(* IEC 61131-3 sources: daoli-st-library/DL_Process (part 27) *)

(* ---- FB_DL_ChillerCondReset.st ---- *)
(*
  FB_DL_ChillerCondReset  —  冷水机组冷凝压力重置（室外湿球联动限幅） / Chiller condensing-pressure setpoint reset driven by outdoor wet-bulb with clamping
  分类 Category : DL_Process
  版本 Version  : 1.0.0
  来源 Source   : t1-2-oscat-building — 楼宇冷站冷凝压力重置族深化
  溯源 Origin   : 道莅 clean-room 实现；湿球联动线性重置 + 死区 + 步长限幅为公开 HVAC 节能控制律，未复制任何源码行
  功能 Function : 1) 目标设定 fCondSpKpa = fWetBulbC × fSlopeKpaPerK + fOffsetKpa；
                  2) 硬限幅钳制到 [fSpMinKpa, fSpMaxKpa]（先限幅后限速，顺序固定）；
                  3) 步长限速：单次调用变化量不超过 fStepMaxKpa（向上与向下同限）；
                  4) 死区保持：|候选 - 当前输出| < fDeadbandKpa 时输出保持不变（避免阀位抖动）；
                  5) 故障级单码 03A3，归因由 eCause 独立成员承载（R190）；
                  6) 信息级 04CB = 重置激活沿（进 eRun 单拍）；7) 解除式全当拍量（R240）。
  接口 Interface: 输入湿球/斜率/偏置/上下限/死区/步长；输出设定值与限幅/限速镜像
  边界 Boundary : ① 组态闸：fSlopeKpaPerK <= 0.0、fSpMaxKpa <= fSpMinKpa、fStepMaxKpa <= 0.0、
                  fDeadbandKpa < 0.0、fWetBulbMaxC <= fWetBulbMinC 任一成立 → 03A3 锁存；
                  ② 湿球非有限（NaN 自反 + Inf 差值自减）或越量程 → 03A3 锁存，输出保持上一有效值
                  （冻结保持，非降级）；③ 浮点判据全容差式，禁 = / <> 判等；
                  ④ 无 TON 跨相复用（仅一个激活沿 R_TRIG + 一个 R_TRIG 复位沿），段 0 无条件调用；
                  ⑤ 故障相迁出唯一路径 = bReset 上升沿；⑥ 零全局耦合（无 GVL / %I %Q %M）。
  依赖 Depends  : Standard.library（R_TRIG）
  码表 Error codes（Process 段 0005，故障窗口 03A3 / 信息窗口 04CB）:
    16#0005_03A3 故障级：冷凝压力重置故障总码（组态非法 / 湿球非有限 / 湿球越量程），
                 锁存至 bReset 上升沿；归因见 eCause，不新增码位（派单硬约束单码）
    16#0005_04CB 信息级：重置激活沿（bEnable 上升进入 eRun 单拍）
  修订历史 Revision :
    2026-11-19  v1.0.0  R43 首版（批次 2 · 序号 7）
*)

TYPE E_DL_CcrState :
(
    eIdle  := 0,      // 未使能：输出冻结上一值 / Idle, output frozen
    eRun   := 10,     // 重置运行中 / Reset active
    eFault := 90      // 故障锁存相 / Fault latched phase
);
END_TYPE

TYPE E_DL_CcrCause :
(
    eNone       := 0, // 无故障成因 / No cause
    eCfgIllegal := 1, // 组态非法 / Illegal configuration
    eWbNonFin   := 2, // 湿球输入非有限 / Wet-bulb non-finite
    eWbRange    := 3  // 湿球越量程 / Wet-bulb out of range
);
END_TYPE

FUNCTION_BLOCK FB_DL_ChillerCondReset
VAR_INPUT
    fWetBulbC      : REAL := 10.0;     // 室外湿球温度 [°C] / Outdoor wet-bulb temperature
    fWetBulbMinC   : REAL := -20.0;    // 湿球量程下限 [°C] / Wet-bulb range low
    fWetBulbMaxC   : REAL := 45.0;     // 湿球量程上限 [°C] / Wet-bulb range high
    fSlopeKpaPerK  : REAL := 2.0;      // 联动斜率 [kPa/K]，域 > 0 / Reset slope
    fOffsetKpa     : REAL := 400.0;    // 联动偏置 [kPa] / Reset offset
    fSpMinKpa      : REAL := 500.0;    // 设定下限 [kPa] / Setpoint low limit
    fSpMaxKpa      : REAL := 900.0;    // 设定上限 [kPa] / Setpoint high limit
    fDeadbandKpa   : REAL := 5.0;      // 死区 [kPa]，域 >= 0 / Deadband
    fStepMaxKpa    : REAL := 10.0;     // 单次限速步长 [kPa]，域 > 0 / Rate limit step
    bEnable        : BOOL := FALSE;    // 重置使能（电平）[-] / Reset enable
    bReset         : BOOL := FALSE;    // 复位命令，上升沿清故障 [-] / Reset edge
END_VAR
VAR_OUTPUT
    eState         : E_DL_CcrState;    // 状态出口，段 6 单点映射 / State outlet
    eCause         : E_DL_CcrCause;    // 故障成因出口（R190） / Fault cause outlet
    fCondSpKpa     : REAL;             // 冷凝压力设定 [kPa] / Condensing pressure setpoint
    bLimited       : BOOL;             // 限幅生效镜像 [-] / Clamp active mirror
    bDbHold        : BOOL;             // 死区保持镜像 [-] / Deadband hold mirror
    bError         : BOOL;             // 故障锁存标志 [-] / Fault latch flag
    nErrId         : UDINT;            // 事件码，0 = 无事件 / Event code
END_VAR
VAR
    _eState        : E_DL_CcrState := E_DL_CcrState.eIdle;   // 内部相位（CASE 唯一写入目标） / Internal phase
    _eCause        : E_DL_CcrCause := E_DL_CcrCause.eNone;   // 故障成因锁存（锁存量） / Latched cause
    rtEnable       : R_TRIG;           // 使能沿实例，每周期无条件调用 / Enable edge
    rtReset        : R_TRIG;           // 复位沿实例，每周期无条件调用 / Reset edge
    _fSp           : REAL;             // 设定输出保持槽（持久） / Setpoint holding slot
    _fRawKpa       : REAL;             // 未限幅原始设定 [kPa]（当拍量） / Raw setpoint
    _fClampKpa     : REAL;             // 限幅后候选 [kPa]（当拍量） / Clamped candidate
    _bClampOn      : BOOL;             // 限幅生效当拍量 [-] / Clamp active
    _bNonFin       : BOOL;             // 湿球非有限当拍量 [-] / Wet-bulb non-finite
    _bRangeBad     : BOOL;             // 湿球越量程当拍量 [-] / Wet-bulb out of range
    _bCfgBad       : BOOL;             // 组态非法当拍量 [-] / Config illegal
    _bFault        : BOOL;             // 故障锁存位（锁存量） / Latched fault bit
    _uFault        : UDINT;            // 故障码锁存（锁存量） / Latched fault code
    _uInfo         : UDINT;            // 信息码，每拍重算 / Transient info code
END_VAR

(* —— 段 0：沿实例无条件周期刷新 + 当拍量判据 —— *)
_fRawKpa := fWetBulbC * fSlopeKpaPerK + fOffsetKpa;                       // 联动原始设定 [kPa] / Raw linked setpoint
_bNonFin := (fWetBulbC <> fWetBulbC) OR ((fWetBulbC - fWetBulbC) <> (fWetBulbC - fWetBulbC));   // NaN/Inf 双判 / NaN and Inf
_bRangeBad := (fWetBulbC < fWetBulbMinC) OR (fWetBulbC > fWetBulbMaxC);    // 量程判据（双侧直比） / Range verdict
_bCfgBad := (fSlopeKpaPerK <= 0.0) OR (fSpMaxKpa <= fSpMinKpa) OR (fStepMaxKpa <= 0.0)
            OR (fDeadbandKpa < 0.0) OR (fWetBulbMaxC <= fWetBulbMinC);     // 组态非法当拍量 / Config illegal
rtEnable(CLK := bEnable);                                                 // 使能沿，每拍必调 / Enable edge
rtReset(CLK := bReset);                                                   // 复位沿，每拍必调 / Reset edge

(* —— 段 1：单拍量预清零（锁存量与设定保持槽不入清单） —— *)
_uInfo := 16#0000_0000;            // 信息码每拍重算 / Info recomputed
bLimited := FALSE;                 // 限幅镜像缺省 FALSE / Clamp mirror default
bDbHold := FALSE;                  // 死区镜像缺省 FALSE / Deadband mirror default
nErrId := 16#0000_0000;            // 事件码缺省无事件 / Event code default

(* —— 段 2：复位沿 + 组态域闸 —— *)
IF rtReset.Q THEN                              // rtReset.Q = 当拍量 / current scan
    _bFault := FALSE;                          // 清故障锁存位（锁存量） / Clear fault latch
    _uFault := 16#0000_0000;                   // 清故障锁存码（锁存量） / Clear fault code
    _eCause := E_DL_CcrCause.eNone;            // 清成因（锁存量） / Clear cause
    IF _eState = E_DL_CcrState.eFault THEN
        _eState := E_DL_CcrState.eIdle;        // 故障相迁出：回未使能 / Fault exit to idle
    END_IF
END_IF
IF _bCfgBad THEN                               // 组态域闸 / Config gate
    _uFault := 16#0005_03A3;                   // 故障级：重置故障总码 / Process fault code
    _eCause := E_DL_CcrCause.eCfgIllegal;      // 归因：组态非法 / Cause: illegal config
    _bFault := TRUE;                           // 标志与码位配对（R45） / Flag paired with code
END_IF

(* —— 段 3：湿球非有限 / 越量程（判据当拍量） —— *)
IF (NOT _bFault) AND _bNonFin THEN             // 非有限锁存 / Non-finite latch
    _uFault := 16#0005_03A3;
    _eCause := E_DL_CcrCause.eWbNonFin;        // 归因：非有限 / Cause: non-finite
    _bFault := TRUE;
END_IF
IF (NOT _bFault) AND (NOT _bNonFin) AND _bRangeBad THEN   // 越量程锁存 / Range latch
    _uFault := 16#0005_03A3;
    _eCause := E_DL_CcrCause.eWbRange;         // 归因：越量程 / Cause: out of range
    _bFault := TRUE;
END_IF

(* —— 段 4：故障解除式（R240；全当拍量）：rtReset.Q / NOT _bCfgBad / NOT _bNonFin / NOT _bRangeBad —— *)
IF rtReset.Q AND (NOT _bCfgBad) AND (NOT _bNonFin) AND (NOT _bRangeBad) THEN
    _bFault := FALSE;                          // 清故障锁存位（锁存量） / Clear fault latch
    _uFault := 16#0000_0000;                   // 清故障锁存码（锁存量） / Clear fault code
    _eCause := E_DL_CcrCause.eNone;            // 清成因（锁存量） / Clear cause
END_IF

(* —— 段 4A：故障锁存相位迁移闸（输出冻结上一有效值，非降级） —— *)
IF _bFault AND (_eState <> E_DL_CcrState.eFault) THEN
    _eState := E_DL_CcrState.eFault;           // 锁存即入故障相 / Latch enters fault phase
END_IF

(* —— 段 5：相位机（CASE 全覆盖 + ELSE 兜底） —— *)
CASE _eState OF

E_DL_CcrState.eIdle:
    IF rtEnable.Q AND (NOT _bFault) THEN       // 使能上升沿启动 / Enable rising starts
        _uInfo := 16#0005_04CB;                // 信息级：重置激活沿 / Info: reset active edge
        _eState := E_DL_CcrState.eRun;         // 进运行相 / Enter run
    END_IF

E_DL_CcrState.eRun:
    IF NOT bEnable THEN                        // 撤使能：回未使能（输出冻结） / Disable returns idle
        _eState := E_DL_CcrState.eIdle;
    ELSE
        _fClampKpa := _fRawKpa;                            // 候选 = 原始设定 / Candidate from raw
        IF _fClampKpa < fSpMinKpa THEN                     // 下限钳制 / Low clamp
            _fClampKpa := fSpMinKpa;
            _bClampOn := TRUE;
        ELSIF _fClampKpa > fSpMaxKpa THEN                  // 上限钳制 / High clamp
            _fClampKpa := fSpMaxKpa;
            _bClampOn := TRUE;
        ELSE
            _bClampOn := FALSE;                            // 未限幅 / No clamp
        END_IF
        IF ABS(_fClampKpa - _fSp) < fDeadbandKpa THEN      // 死区内保持（容差式比较） / Deadband hold
            bDbHold := TRUE;
        ELSIF (_fClampKpa - _fSp) > fStepMaxKpa THEN       // 向上限速 / Upward rate limit
            _fSp := _fSp + fStepMaxKpa;
        ELSIF (_fSp - _fClampKpa) > fStepMaxKpa THEN       // 向下限速 / Downward rate limit
            _fSp := _fSp - fStepMaxKpa;
        ELSE
            _fSp := _fClampKpa;                            // 直接跟随 / Direct follow
        END_IF
        IF (_fSp < fSpMinKpa) THEN                         // 限速后二次下限复核 / Post-limit low check
            _fSp := fSpMinKpa;
        ELSIF (_fSp > fSpMaxKpa) THEN                      // 限速后二次上限复核 / Post-limit high check
            _fSp := fSpMaxKpa;
        END_IF
    END_IF

E_DL_CcrState.eFault:
    ;                                          // 故障相：输出冻结，仅段 4 复位沿可迁出 / Frozen, reset only

ELSE
    _uFault := 16#0005_03A3;                   // 故障级：非法相位兜底（归并总码） / Illegal phase fallback
    _eCause := E_DL_CcrCause.eCfgIllegal;      // 归因：相位非法归并组态 / Cause: phase illegal
    _bFault := TRUE;
    _eState := E_DL_CcrState.eFault;           // 强制回故障相 / Force fault phase

END_CASE

(* —— 段 6：出口单点映射（名实同源；锁存码回放） —— *)
fCondSpKpa := _fSp;                            // 设定值出口 / Setpoint outlet
bLimited := _bClampOn AND (NOT _bFault);       // 限幅镜像 / Clamp mirror
bDbHold := bDbHold AND (NOT _bFault);          // 死区保持镜像 / Deadband mirror
IF _bFault THEN
    nErrId := _uFault;                         // 故障锁存码回放 / Replay latched code
ELSE
    nErrId := _uInfo;                          // 信息码 / Transient info
END_IF
bError := _bFault;                             // 故障标志同源 / Flag from latch
eState := _eState;                             // 状态出口 / State outlet
eCause := _eCause;                             // 成因出口 / Cause outlet

END_FUNCTION_BLOCK

(* ---- FB_DL_ChillerDoorPurgeSeq.st ---- *)
(*
    FB_DL_ChillerDoorPurgeSeq —— 冷机检修门吹扫联锁时序
    ------------------------------------------------------------------
    分类      : DL_Process / Interlock
    前缀      : FB_DL_
    版本      : 1.0.0
    溯源      : clean-room 自有实现；仅借鉴「先吹扫置换、后放行开门」的受限空间
                进入公开安全常识语义，未复制任何闭源厂商源码，码位 100% 自有
    平台      : 纯 IEC 61131-3，CODESYS V3.5+ / TwinCAT 3 / InoProShop / Machine Expert 通用
    作者      : 道莅代码库 · PLC编程专家（R76 冲刺批 C3 · #3）
    ------------------------------------------------------------------
    功能说明  : 冷机检修门「吹扫联锁」唯一时序属主件：门关到位确认 → 风压建立确认
                （fAirPress > fPressMin 持续 tPressQual，超 tPressTo 未建立报 1F00）
                → 吹扫倒计时（tPurgeDur）→ 吹扫完成（bDone 单拍脉冲）→ 放行门开允许
                （bDoorPermit）。任一异常（门中途打开 / 风压跌落 / 确认超时）→
                回退安全态（吹扫输出与开门允许同时撤销）并锁存故障，须 bReset 复位；
                bEStop 急停为最高优先，任意态立即回安全态并锁存 1F03。
                边界：只产出吹扫输出与开门允许，不驱动门电机、不判冷剂浓度。
    序列      : eIdle --bDoorClosed--> ePressQual --fbPressQual.Q--> ePurging
                --fbPurge.Q--> eReady（bDoorPermit）--门正常打开--> eIdle；
                ePressQual/ePurging --门中途打开--> eFault（1F02）；
                ePurging --风压跌落--> eFault（1F01）；ePressQual --超时--> eFault（1F00）。
    错误码    : 16#0005_1F00 风压建立确认超时（tPressTo 内未持续达标）——故障级
                16#0005_1F01 吹扫期间风压跌落（低于 fPressMin）——故障级
                16#0005_1F02 门中途打开（风压确认或吹扫中）——故障级
                16#0005_1F03 急停触发——故障级，最高优先，任意态立即安全态
                16#0005_1F04 参数/采样非法（fAirPress 非有限 / 阈值非正 / 时间为零）——故障级
                16#0005_1F05 CASE 落 ELSE 兜底——故障级
    码位总账  : 16#0005_1F00..1F05 全部定义并使用，无空悬码位
    状态机    : E_DL_PurgeState（eIdle / ePressQual / ePurging / eReady / eFault），
                CASE 含 ELSE 兜底：落 ELSE 置 16#0005_1F05、回安全态转 eFault。
                全部故障码锁存至复位沿：bReset 上升沿且 bEStop 已解除方可复位；
                吹扫完成脉冲 bDone 为单拍位：内部 _bDonePulse 置位 → 统一出口
                映射单拍发布（两段式，防同拍抹除）。
    安全优先级: 段 3 急停拦截在参数门禁与状态机之前执行，任意态（含 eFault）急停
                即重锁存 1F03 并保持安全态输出；安全态 = 吹扫输出 OFF + 开门允许 OFF。
    定时器    : 三只 TON + 两只 R_TRIG 在本体段 1 无条件周期刷新（R7），绝不放入
                CASE/IF，实例无跨相复用。
    防御口径  : 浮点比较一律阈值比较（禁 =/<>）；本件无除法运算；非有限判定按
                NaN f<>f、±Inf (f-f)<>(f-f)。
    修订记录  : 2026-11-23 v1.0.0 首次入库（R76 冲刺批 C3 · #3）
*)
TYPE E_DL_PurgeState :
(
    eIdle       := 0,   // 待机，等门关到位，吹扫与放行全撤销 / idle, waiting for the closed door, purge and permit both off
    ePressQual  := 10,  // 风压建立确认中，fAirPress 持续达标计时 / pressure qualifying, timing while air pressure stays above the minimum
    ePurging    := 20,  // 吹扫倒计时中，风压须持续保持 / purging, countdown running while pressure must hold
    eReady      := 30,  // 吹扫完成，开门允许放行 / purge complete, door-open permit granted
    eFault      := 40   // 故障，安全态保持，故障码锁存至复位沿 / fault, safe state held, code latched until the reset edge
);
END_TYPE

FUNCTION_BLOCK FB_DL_ChillerDoorPurgeSeq
VAR_INPUT
    bDoorClosed : BOOL;                  // 门关到位反馈，TRUE = 已关严 / door closed feedback, TRUE = fully closed
    fAirPress   : REAL;                  // 吹扫风压采样 [kPa] / purge air pressure sample [kPa]
    fPressMin   : REAL := 5.0;           // 风压建立阈值 [kPa]，必须大于 0 / pressure qualification threshold [kPa], must exceed zero
    tPressQual  : TIME := T#1S;          // 风压确认持续时间 [ms]，必须大于 0 / pressure qualification dwell [ms], must exceed zero
    tPressTo    : TIME := T#5S;          // 风压建立超时窗 [ms]，须大于 tPressQual / pressure establish timeout [ms], must exceed tPressQual
    tPurgeDur   : TIME := T#30S;         // 吹扫倒计时时长 [ms]，必须大于 0 / purge duration [ms], must exceed zero
    bEStop      : BOOL;                  // 急停输入，TRUE = 急停，最高优先 / emergency stop, TRUE = stopped, highest priority
    bReset      : BOOL;                  // 故障复位请求，上升沿生效且须急停已解除 / fault reset request, edge-active and requires estop cleared
END_VAR
VAR_OUTPUT
    bPurgeCmd   : BOOL;                  // 吹扫风机/风阀输出，仅确认与吹扫相置位 / purge blower or valve output, asserted in the qualify and purge phases only
    bDoorPermit : BOOL;                  // 门开允许，仅吹扫完成相置位 / door-open permit, asserted in the ready phase only
    bDone       : BOOL;                  // 吹扫完成单拍脉冲，发布后自清 / purge-complete one-scan pulse, self-cleared after publishing
    eState      : E_DL_PurgeState;       // 当前状态镜像输出 / current state mirror output
    nErrCode    : UDINT;                 // 错误码，0 = 无错；故障级码全部锁存回放 / error code, 0 = none; all fault-class codes latched and replayed
    bError      : BOOL;                  // 故障级标志，仅故障级码置位 / fault-class flag, raised only by fault-class codes
    bValid      : BOOL;                  // 输出可用标志，= NOT bError / outputs valid flag, equals NOT bError
END_VAR
VAR
    fbPressQual : TON;                   // 风压确认定时器，仅 ePressQual 使用 / pressure qualification timer, ePressQual only
    fbPressTo   : TON;                   // 风压建立超时定时器，仅 ePressQual 使用 / pressure establish timeout timer, ePressQual only
    fbPurge     : TON;                   // 吹扫倒计时定时器，仅 ePurging 使用 / purge countdown timer, ePurging only
    rtReset     : R_TRIG;                // 复位上升沿检测 / reset rising-edge detector
    _eState     : E_DL_PurgeState;       // 当前状态 / current state
    _uErrLatch  : UDINT;                 // 故障码锁存副本，故障态每拍回放 / latched fault code republished inside the fault state
    _bDonePulse : BOOL;                  // 完成脉冲源，段 2 发布后立刻自清 / completion pulse source, published then cleared in segment 2
    _bGateOk    : BOOL;                  // 参数与采样门禁结果 / parameter and sample gate result
END_VAR
VAR CONSTANT
    DL_CDP_ZERO : REAL := 0.0;           // 零值常量，避免裸字面量 [kPa] / zero constant avoiding a bare literal [kPa]
    DL_CDP_T_ZERO : TIME := T#0S;        // 零时间常量，参数门禁用 / zero time constant for the parameter gate
END_VAR

// 段 1｜定时器与边缘检测无条件周期刷新（R7：严禁放入 IF / CASE，实例无跨相复用）
// segment 1, timers and edge detectors refreshed unconditionally, never inside IF/CASE, no cross-phase reuse
fbPressQual(IN := (_eState = E_DL_PurgeState.ePressQual) AND (fAirPress > fPressMin) AND _bGateOk, PT := tPressQual);
fbPressTo(IN := (_eState = E_DL_PurgeState.ePressQual), PT := tPressTo);
fbPurge(IN := (_eState = E_DL_PurgeState.ePurging), PT := tPurgeDur);
rtReset(CLK := bReset);

// 段 2｜输出与错误状态预置；故障态从锁存副本回放；完成脉冲统一出口单拍发布（两段式）
// segment 2, preset outputs and error status; the fault state replays from the latch; the done pulse is published one scan via the unified exit
bDone := _bDonePulse;                    // 发布上一拍置的完成脉冲 / publish the pulse latched last scan
_bDonePulse := FALSE;                    // 发布即自清，保证只出现一拍 / clear right after publishing so the pulse lasts one scan
nErrCode := 0;                           // 预置无错误码 / preset no error code
bError := FALSE;                         // 预置无故障标志 / preset no fault flag
bValid := TRUE;                          // 预置输出可用 / preset outputs valid
IF _eState = E_DL_PurgeState.eFault THEN
    nErrCode := _uErrLatch;              // 重发布锁存故障码，HMI 不会看到码位闪断 / republish the latched fault code
    bError := TRUE;                      // 故障态恒置故障标志 / fault flag stays raised in the fault state
    bValid := FALSE;                     // 故障态输出不可信 / outputs not valid in the fault state
END_IF

// 段 3｜急停最高优先拦截 + 参数/采样门禁：急停任意态立即锁存 1F03 回安全态；
//        门禁非法锁存 1F04 转故障；已在故障态不覆盖原锁存码
// segment 3, estop has the highest priority and latches 1F03 from any state including fault;
//        the parameter gate latches 1F04; an existing latch inside the fault state is not overwritten
IF bEStop THEN
    _uErrLatch := 16#0005_1F03;          // 锁存急停码（任意态含 eFault 均可覆盖更新）/ latch the estop code, overridable from any state
    nErrCode := 16#0005_1F03;            // 故障级码赋值 3 行内置 bError / fault-class assignment with bError inline
    bError := TRUE;
    bValid := FALSE;
    _eState := E_DL_PurgeState.eFault;   // 立即回安全态，本拍 CASE 按 eFault 分派 / jump to the safe state, CASE dispatches on eFault
ELSE
    _bGateOk := (fPressMin > DL_CDP_ZERO) AND (tPressQual > DL_CDP_T_ZERO)
            AND (tPressTo > DL_CDP_T_ZERO) AND (tPurgeDur > DL_CDP_T_ZERO)
            AND (tPressTo > tPressQual);
    IF (fAirPress <> fAirPress) OR ((fAirPress - fAirPress) <> (fAirPress - fAirPress)) THEN
        _bGateOk := FALSE;               // 风压采样 NaN 或 ±Inf，非有限判定 / pressure sample NaN or infinite
    END_IF
    IF (NOT _bGateOk) AND (_eState <> E_DL_PurgeState.eFault) THEN
        _uErrLatch := 16#0005_1F04;      // 锁存参数/采样非法码 / latch the illegal parameter or sample code
        nErrCode := 16#0005_1F04;        // 故障级码赋值 3 行内置 bError / fault-class assignment with bError inline
        bError := TRUE;
        bValid := FALSE;
        _eState := E_DL_PurgeState.eFault; // 参数不可信直接转故障 / untrusted parameters jump to fault
    END_IF
END_IF

// 段 4｜主状态机：CASE + ELSE 兜底（R6）；每个相注明 拍 N 进入 / 本拍行为 / 拍 N+1 转出
// segment 4, main state machine, CASE with ELSE fallback; each phase notes entry, per-scan behaviour and exits
CASE _eState OF
E_DL_PurgeState.eIdle:
    // 拍 N 进入：复位后或门正常打开后；本拍行为：全撤销等待；拍 N+1 转出：门关到位 → ePressQual
    // entered after reset or a normal door opening; everything off while waiting; exits to ePressQual on the closed door
    IF bDoorClosed AND _bGateOk THEN
        _eState := E_DL_PurgeState.ePressQual; // 进风压确认相，下一拍计时启动 / enter pressure qualification, timing starts next scan
    END_IF

E_DL_PurgeState.ePressQual:
    // 拍 N 进入：门关到位；本拍行为：风压达标则 fbPressQual 计时；拍 N+1 转出四路：
    // 计时到 → ePurging；门中途打开 → eFault（1F02）；确认超时 → eFault（1F00）；门禁 → eFault（段 3）
    // entered on the closed door; timer runs while pressure holds; exits to ePurging on Q,
    // to eFault on a mid-sequence door opening (1F02) or on the establish timeout (1F00)
    IF NOT bDoorClosed THEN
        _uErrLatch := 16#0005_1F02;      // 锁存门中途打开码 / latch the mid-sequence door opening code
        nErrCode := 16#0005_1F02;        // 故障级码赋值 3 行内置 bError / fault-class assignment with bError inline
        bError := TRUE;
        bValid := FALSE;
        _eState := E_DL_PurgeState.eFault; // 回安全态，吹扫与放行同拍撤销 / safe state, purge and permit drop the same scan
    ELSIF fbPressQual.Q THEN
        _eState := E_DL_PurgeState.ePurging; // 风压确认通过，进吹扫倒计时 / pressure qualified, start the purge countdown
    ELSIF fbPressTo.Q THEN
        _uErrLatch := 16#0005_1F00;      // 锁存风压建立超时码 / latch the pressure establish timeout code
        nErrCode := 16#0005_1F00;        // 故障级码赋值 3 行内置 bError / fault-class assignment with bError inline
        bError := TRUE;
        bValid := FALSE;
        _eState := E_DL_PurgeState.eFault; // 超时回退安全态 / roll back to the safe state on timeout
    END_IF

E_DL_PurgeState.ePurging:
    // 拍 N 进入：风压确认通过；本拍行为：吹扫输出保持、倒计时走、风压须持续达标；
    // 拍 N+1 转出三路：倒计时到 → eReady（置完成脉冲源）；风压跌落 → eFault（1F01）；
    // 门中途打开 → eFault（1F02）
    // entered after qualification; purge output held, countdown running, pressure must hold;
    // exits to eReady with the pulse source on Q, to eFault on pressure drop (1F01) or door opening (1F02)
    IF NOT bDoorClosed THEN
        _uErrLatch := 16#0005_1F02;      // 锁存门中途打开码 / latch the mid-sequence door opening code
        nErrCode := 16#0005_1F02;        // 故障级码赋值 3 行内置 bError / fault-class assignment with bError inline
        bError := TRUE;
        bValid := FALSE;
        _eState := E_DL_PurgeState.eFault; // 回安全态 / return to the safe state
    ELSIF fAirPress < fPressMin THEN
        _uErrLatch := 16#0005_1F01;      // 锁存风压跌落码 / latch the pressure drop code
        nErrCode := 16#0005_1F01;        // 故障级码赋值 3 行内置 bError / fault-class assignment with bError inline
        bError := TRUE;
        bValid := FALSE;
        _eState := E_DL_PurgeState.eFault; // 风压跌落立即回退 / roll back at once on the pressure drop
    ELSIF fbPurge.Q THEN
        _bDonePulse := TRUE;             // 置完成脉冲源，段 2 统一出口单拍发布 / set the pulse source, published one scan via segment 2
        _eState := E_DL_PurgeState.eReady;   // 吹扫完成，进放行相 / purge complete, enter the ready phase
    END_IF

E_DL_PurgeState.eReady:
    // 拍 N 进入：吹扫倒计时到；本拍行为：开门允许置位（输出映射段）、吹扫输出撤销；
    // 拍 N+1 转出：门正常打开（关反馈消失）→ eIdle，下次关门重新吹扫
    // entered when the countdown elapsed; permit asserted via the output map while the purge output drops;
    // exits to eIdle when the door actually opens, the next closure restarts the purge
    IF NOT bDoorClosed THEN
        _eState := E_DL_PurgeState.eIdle;    // 门已开，正常返回待机 / door opened, normal return to idle
    END_IF

E_DL_PurgeState.eFault:
    // 拍 N 进入：任一故障级路径；本拍行为：安全态保持、锁存码回放；拍 N+1 转出：
    // bReset 上升沿且急停已解除 → eIdle（门关反馈丢失自动回 eIdle 等下次关门）
    // entered from any fault path; safe state held and the latch replays; exits to eIdle only on
    // a reset edge with the estop cleared
    IF rtReset.Q AND (NOT bEStop) THEN
        _uErrLatch := 0;                 // 清锁存码 / clear the latched code
        _eState := E_DL_PurgeState.eIdle;    // 回待机，等下次门关到位 / back to idle for the next closure
    END_IF

ELSE
    // 非法状态拦截：任何未定义枚举值一律锁存兜底码并转故障（R6）
    // illegal-state interception, any undefined enum value latches the fallback code and goes to fault
    _uErrLatch := 16#0005_1F05;          // 锁存兜底码 / latch the fallback code
    nErrCode := 16#0005_1F05;            // 故障级码赋值 3 行内置 bError / fault-class assignment with bError inline
    bError := TRUE;
    bValid := FALSE;
    _eState := E_DL_PurgeState.eFault;
END_CASE

// 段 5｜输出映射：吹扫输出仅确认/吹扫相保持，开门允许仅就绪相置位，其余一律撤销（双保险）
// segment 5, output map; purge output held only in qualify/purge, permit only in ready, everything else dropped as a double cut
bPurgeCmd := (_eState = E_DL_PurgeState.ePressQual)
          OR (_eState = E_DL_PurgeState.ePurging);   // 吹扫输出按相映射 / purge output mapped by phase
bDoorPermit := (_eState = E_DL_PurgeState.eReady);   // 开门允许仅在放行相 / permit only in the ready phase
eState := _eState;                                   // 状态镜像输出 / state mirror output

END_FUNCTION_BLOCK

(* ---- FB_DL_ChillerLiftOptimize.st ---- *)
(*
  Component : FB_DL_ChillerLiftOptimize
  Category  : DL_Process
  Type      : FB
  Version   : 1.0.0
  CodeSeg   : 16#06_0_37
  Summary   : 冷机 Lift（冷凝-蒸发温差）优化限值：温差基线统计窗 + 设定值 RateLimiter 限速输出。
              Chiller lift optimization: condenser-evaporator baseline statistics window plus rate-limited setpoint.
  溯源声明  : 道莅自研 clean-room
  边界安全  : 温度非有限（NaN 自反 + Inf 上限）拦截；基线统计窗点数域闸（≥ 1）；
              统计窗未满时输出冻结在当前值并置 bBaselineReady=FALSE（按派单要点）；
              设定值输出过 RateLimiter 限速（每拍步进钳制，防设定值跳变）；全浮点比较带 fEps 容差。
  复用      : 无
*)

FUNCTION_BLOCK FB_DL_ChillerLiftOptimize
VAR_INPUT
    bRun        : BOOL;                 (* 优化使能 · Enable *)
    fCondTC     : LREAL;                (* 冷凝器温度 [degC] · Condenser temperature *)
    fEvapTC     : LREAL;                (* 蒸发器温度 [degC] · Evaporator temperature *)
    nWinScans   : INT := 600;           (* 基线统计窗长 [拍] · Baseline window length *)
    fStepMaxK   : LREAL := 0.1;         (* 设定值每拍最大步进 [K] · Setpoint max step per scan *)
    fDeadK      : LREAL := 0.5;         (* 优化死区 [K]，防频繁调节 · Optimization deadband *)
    fEps        : LREAL := 1.0E-6;      (* 浮点判零容差 [实数域] · Floating zero tolerance *)
END_VAR
VAR_OUTPUT
    fLiftNowK   : LREAL;                (* 当前 Lift [K] · Current lift *)
    fLiftBaseK  : LREAL;                (* 基线平均 Lift [K] · Baseline mean lift *)
    fSetK       : LREAL;                (* 优化设定值输出 [K]，已限速 · Rate-limited setpoint *)
    bBaselineReady: BOOL;               (* 基线窗满标志 · Baseline ready flag *)
    bError      : BOOL;                 (* 故障标志，与故障码配对 · Fault flag paired with codes *)
    uErrorId    : UDINT;                (* 事件码 16#0000_0037，0 无事件 · Event code *)
END_VAR
VAR
    uCode   : WORD;     (* 码位暂存，每拍重算 [码] · Code staging *)
    bSigOk  : BOOL;     (* 输入有效标志 · Input validity flag *)
    fSumK   : LREAL;    (* 窗内 Lift 累加和 [K·拍] · Window sum *)
    nFill   : INT;      (* 窗内已累计拍数 [拍] · Window filled scans *)
    fTargetK: LREAL;    (* 目标设定值 [K] · Target setpoint *)
    fStepK  : LREAL;    (* 本拍实际步进 [K] · Actual step this scan *)
    nCycles : UDINT;    (* 有效拍计数 [拍]，防回卷 · Valid scan count *)
END_VAR
VAR CONSTANT
    DL_CLO_WRAP : UDINT := 4294967290;  (* 计数防回卷余量 [拍] · Counter wrap guard *)
END_VAR

(* === 段 0 · 实例刷新 === *)
(* 无 TON/R_TRIG 实例：基线窗按拍计数；No timer instances, scan-counted window *)

(* === 段 1 · 输入校验与量程闸 === *)
uCode := 16#0000;                       // 每拍清码（可达清零基线）/ Clear codes each scan
bSigOk := (fCondTC = fCondTC) AND (fEvapTC = fEvapTC)               // 非有限拦截 / Non-finite guard
          AND (ABS(fCondTC) < 1.0E308) AND (ABS(fEvapTC) < 1.0E308) // Inf 上限判据 / Inf limit
          AND (nWinScans >= 1)                                      // 窗长域闸 / Window length gate
          AND (fStepMaxK > 0.0) AND (fDeadK >= 0.0);                // 步进正域闸 / Step and deadband gates
IF NOT bSigOk THEN
    uCode := 16#0037;                   // 故障级：域外，输出冻结 / Fault: domain invalid, frozen
END_IF

(* === 段 2 · 主逻辑：Lift 基线统计与设定值限速 === *)
IF bSigOk THEN
    fLiftNowK := fCondTC - fEvapTC;     (* 当前 Lift [K] / Current lift *)
    IF bRun THEN
        IF nFill < nWinScans THEN
            fSumK := fSumK + fLiftNowK; (* 窗内累加 / Accumulate in window *)
            nFill := nFill + 1;         (* 窗计数推进 / Advance the window count *)
            bBaselineReady := FALSE;    (* 窗未满：基线未就绪 / Window not full *)
        ELSE
            fLiftBaseK := fSumK / UDINT_TO_LREAL(INT_TO_UDINT(nWinScans));  (* 基线均值 [K] / Baseline mean *)
            bBaselineReady := TRUE;     (* 窗满：基线就绪 / Window full, baseline ready *)
            IF fLiftNowK > (fLiftBaseK + fDeadK) THEN
                fTargetK := fLiftBaseK; (* 超死区回基线目标 / Target back to baseline *)
            ELSE
                fTargetK := fSetK;      (* 死区内保持现值 / Hold inside the deadband *)
            END_IF
        END_IF
    ELSE
        nFill := 0;                     (* 撤使能重开统计窗 / Restart the window on disable *)
        fSumK := 0.0;
        bBaselineReady := FALSE;        (* 撤使能基线失效 / Baseline not ready *)
    END_IF
    (* RateLimiter：设定值每拍步进钳制 / Rate limiter: clamp the per-scan step *)
    fStepK := fTargetK - fSetK;         (* 目标差 [K] / Gap to target *)
    IF fStepK > fStepMaxK THEN
        fSetK := fSetK + fStepMaxK;     (* 正向限速 / Positive rate limit *)
    ELSIF fStepK < (-fStepMaxK) THEN
        fSetK := fSetK - fStepMaxK;     (* 负向限速 / Negative rate limit *)
    ELSE
        fSetK := fTargetK;              (* 一步到位 / Settle to target *)
    END_IF
END_IF

(* === 段 3 · 输出映射与故障码 === *)
IF bSigOk THEN
    IF nCycles < DL_CLO_WRAP THEN
        nCycles := nCycles + 1;         (* 有效拍计数 / Count valid scans *)
    END_IF
END_IF
bError := (uCode <> 16#0000);           (* 故障标志配对 / Fault flag paired *)
uErrorId := WORD_TO_UDINT(uCode);       (* 码位单点写入（16#0000_0037 形态）/ Single write point *)
END_FUNCTION_BLOCK

(* ---- FB_DL_ChillerSeqMgr.st ---- *)
//==============================================================================
// 功能块：FB_DL_ChillerSeqMgr ｜ 中文名称：冷水机组群控调度
// 所属子库：DL_Process ｜ 版本：v1.0.0 ｜ 兼容：CODESYS V3.5+ / TwinCAT 3 / 汇川 InoProShop
// 功能描述：6 台冷水机组群控：按平滑后负荷率加减机（加/减各带独立延迟，双延迟防抖动）
//           + 主备轮值均衡（委托 FB_DL_DutyStandbyRotation，最短运行/最短停机时长逻辑
//           一律由该件承担，本件只把 tMinRun/tMinStop 转发，绝不重复实现）+ 故障切备
//           （故障台由轮值件跳过）+ 供水低温保护（强制减机，防冻管）。本件不内联机组建模
//           与机组自身控制（压缩机/冷却水阀/防冻判据归设备层），只出启停命令与调度诊断。
// 开源溯源 (Origin)：道莅原创实现（参考 公开工程惯例 分类与参数域）
// 单位表：温度[摄氏度] / 负荷率与阈值[百分数] / 延迟与最小时长[min] / 扫描间隔[ms] /
//         台数[台] / 机组号[号]
// 错误码表：16#0005_040C 信息级（加/减机延迟计时中，尚未动作，不置 bError）/
//           16#0005_040D 信息级（供水温度低限保护强制减机，信息级不锁故障但强制动作）/
//           16#0005_0354 故障级（无可用机组：全故障或全不就绪，工艺停机级，置 bError）/
//           16#0005_0355 故障级（负荷率/阈值组态非法：减机阈值 ≥ 加机阈值、阈值越
//           0~100、台数组态非法；兼轮值件参数冲突透传——轮值件 bError 透传复位且只在
//           故障相处置，R115）/ 16#0005_0356 故障级（输入非有限独立分支显式映射入本槽，
//           兼状态机 ELSE 非法状态兜底）。0356 共用反证句：非有限与非法状态在现有输出
//           组合下不可观测出差异（均为 bError + 全撤指令 + bValid 撤 + eState 进 eFault），
//           §3 未给本件独立非有限槽，故显式复用不越段。
// 状态机：E_DL_ChillerGroupState（eIdle=0 待机 / eRunning=10 稳态调度 /
//           eStageUp=20 加机延迟中 / eStageDown=30 减机延迟中 / eLowSupply=40 供水低温
//           保护 / eFault=99 故障兜底），CASE 含 ELSE 兜底，ELSE 置 0356 且全撤指令。
// 边界行为：① 无可用机组（全故障或全不就绪）→ 故障 0354 + bNoAvailable（工艺停机级，
//           非提示级）；② 阈值组态非法（减机阈值 ≥ 加机阈值、阈值不在 0~100）→ 故障
//           0355；③ 供水温度 < fSupplyLowC → 强制减机一台 + 信息 040D + bLowSupplyProtect
//           （防冻管，信息级不锁故障但强制动作）；④ 加减机延迟计时中 → 信息 040C；
//           ⑤ 需求台数域 0~6 钳位，且不超过可用台数；⑥ 非有限 → 独立分支显式置 0356，
//           全撤指令；⑦ 失能 → 全撤指令 + bValid := FALSE（R72）；⑧ 轮值调用
//           FB_DL_DutyStandbyRotation（组合调用），tMinRunTime/tMinStopTime 由本件引脚
//           转发，最短运行/停机逻辑不重复实现；轮值件 bError 透传复位并在故障相处置。
// 修订历史：v1.0.0 2026-11-17 首版（R25 派单 · §4.18，依赖 DL_Base 件 FB_DL_DutyStandbyRotation 语义）
//==============================================================================
(*------------------------------------------------------------------------------
 * 枚举: E_DL_ChillerGroupState（归属 DL_Process，与 FB_DL_ChillerSeqMgr 同文件）
 *----------------------------------------------------------------------------*)
TYPE E_DL_ChillerGroupState :
(
    eIdle      := 0,   // 待机：失能，指令全撤 / Idle, all commands dropped
    eRunning   := 10,  // 稳态调度：负荷在双阈值之间 / Steady scheduling, load inside both thresholds
    eStageUp   := 20,  // 加机延迟中：负荷高于加机阈值，等延迟到点 / Stage-up delay running
    eStageDown := 30,  // 减机延迟中：负荷低于减机阈值，等延迟到点 / Stage-down delay running
    eLowSupply := 40,  // 供水低温保护：强制减机 / Supply low-temperature protection, forced stage-down
    eFault     := 99   // 故障兜底：无可用机组/组态非法/非有限/非法状态 / Fault fallback
);
END_TYPE

(*==============================================================================
 * 功能块: FB_DL_ChillerSeqMgr
 * 调用约定: 每个扫描周期无条件调用一次；uDeltaTimeMs 必须注入真实任务间隔。
 *============================================================================*)
FUNCTION_BLOCK FB_DL_ChillerSeqMgr
VAR_INPUT
    abChillerReady   : ARRAY[0..5] OF BOOL;        // 机组就绪（无故障、无就地、无禁止）/ Unit ready
    abChillerRunning : ARRAY[0..5] OF BOOL;        // 机组运行反馈 / Unit running feedback
    abChillerFault   : ARRAY[0..5] OF BOOL;        // 机组故障（轮值件跳过并允许立即停机）/ Unit fault
    fSupplyC         : LREAL;                      // 冷冻水供水温度 [摄氏度] / Chilled-water supply temperature [degC]
    fReturnC         : LREAL;                      // 冷冻水回水温度 [摄氏度] / Chilled-water return temperature [degC]
    fLoadPct         : LREAL;                      // 当前负荷率 [百分数] / Current load [percent]
    fStageUpThrPct   : LREAL := 85.0;              // 加机阈值 [百分数] / Stage-up threshold [percent]
    fStageDownThrPct : LREAL := 40.0;              // 减机阈值 [百分数] / Stage-down threshold [percent]
    tStageUpDelay    : TIME := T#10M;              // 加机延迟 [min] / Stage-up delay [min]
    tStageDownDelay  : TIME := T#15M;              // 减机延迟 [min] / Stage-down delay [min]
    tMinRun          : TIME := T#15M;              // 最小运行时长 [min]，转发轮值件 / Minimum run time, forwarded
    tMinStop         : TIME := T#10M;              // 最小停机时长 [min]，转发轮值件 / Minimum stop time, forwarded
    fSupplyLowC      : LREAL := 4.0;               // 供水低温保护门限 [摄氏度] / Supply low-temperature threshold [degC]
    bEnable          : BOOL;                       // 总使能 / Master enable
    bReset           : BOOL;                       // 复位，上升沿清调度状态并透传轮值件 / Reset, rising edge clears the schedule and the duty block
    uDeltaTimeMs     : UDINT;                      // 扫描间隔 [ms]，调用方注入，禁系统时间函数 / Scan interval [ms], caller-injected
END_VAR
VAR_OUTPUT
    abStartCmd       : ARRAY[0..5] OF BOOL;        // 机组启停命令（FALSE = 停）/ Unit start command, FALSE = stop
    nLeadChiller     : INT;                        // 领机号 0~5，-1 = 无 / Lead chiller 0..5, -1 = none
    nRunningCmd      : INT;                        // 指令开机台数 [台] / Commanded running units [pcs]
    fLoadAvgPct      : LREAL;                      // 平滑后负荷率 [百分数] / Smoothed load [percent]
    bStageUpPending  : BOOL;                       // 加机延迟计时中 / Stage-up delay running
    bStageDownPending : BOOL;                      // 减机延迟计时中 / Stage-down delay running
    bNoAvailable     : BOOL;                       // 无可用机组标志 / No available unit flag
    bLowSupplyProtect : BOOL;                      // 供水低温保护生效 / Supply low-temperature protection active
    eErr             : UDINT;                      // 错误码，0 = 无错，码位 16#0005_040C 起信息级、16#0005_0354 起故障级（分带见错误码表） / Error code, 0 = no error, band info/fault per the code table
    bError           : BOOL;                       // 故障级标志，仅故障级错误置位 / Fault-class flag, set only on fault-level codes
    bValid           : BOOL;                       // 命令输出可用标志，失能/故障闸显式 FALSE / Command usable flag, explicit FALSE on disable/fault gates
    eState           : E_DL_ChillerGroupState;     // 主状态机当前状态 / Current state of the main state machine
END_VAR
VAR
    fbReset          : R_TRIG;                     // 复位上升沿检测实例 / Reset rising edge detector
    fbTonUp          : TON;                        // 加机延迟定时器实例 / Stage-up delay timer
    fbTonDown        : TON;                        // 减机延迟定时器实例 / Stage-down delay timer
    fbDuty           : FB_DL_DutyStandbyRotation;  // 主备轮值调度组合实例（DL_Base，契约见手册）/ Duty rotation composed instance
    abUnitReady      : ARRAY[0..7] OF BOOL;        // 轮值件就绪入参（0~5 机组，6~7 空槽）/ Ready input for the duty block
    abUnitRunning    : ARRAY[0..7] OF BOOL;        // 轮值件运行入参（0~5 机组，6~7 空槽）/ Running input for the duty block
    abUnitFault      : ARRAY[0..7] OF BOOL;        // 轮值件故障入参（0~5 机组，6~7 空槽）/ Fault input for the duty block
    abStartCmdDuty   : ARRAY[0..7] OF BOOL;        // 轮值件启停命令暂存（0~5 有效）[—] / Duty start commands staged
    nLeadStage       : INT;                        // 轮值件领机号暂存 [号] / Lead unit staged from the duty block
    bDutyFault       : BOOL;                       // 轮值件故障标志暂存 / Duty fault flag staged
    nDemand          : INT;                        // 需求运行台数（本拍生效值，下一拍送轮值件）[台] / Demand, effective next scan
    nUsable          : INT;                        // 可用机组数 [台] / Usable unit count
    nLoop            : INT;                        // 循环索引 [—] / Loop index
    uGateCode        : UDINT;                      // 机构闸故障码暂存 / Gate fault code staging
    fDtSec           : LREAL;                      // 扫描间隔换算成秒 [s] / Scan interval in seconds [s]
    fAlpha           : LREAL;                      // 负荷率一阶滤波系数 [—] / First-order filter coefficient
    fDenomSec        : LREAL;                      // 滤波系数分母 [s] / Filter denominator [s]
    bNonFin          : BOOL;                       // 非有限判定中间标志 / Non-finite detection intermediate flag
    bNeedUp          : BOOL;                       // 加机需求（瞬时）/ Stage-up need, instantaneous
    bNeedDown        : BOOL;                       // 减机需求（瞬时）/ Stage-down need, instantaneous
    bRearmUp         : BOOL;                       // 加机定时器重装脉冲 / Stage-up timer re-arm pulse
    bRearmDown       : BOOL;                       // 减机定时器重装脉冲 / Stage-down timer re-arm pulse
    bLowSupply       : BOOL;                       // 供水低温判据（瞬时）/ Low supply predicate
    bFirstScan       : BOOL := TRUE;               // 上电首拍标志 / First-scan flag
END_VAR
VAR CONSTANT
    DL_CSM_CODE_INFO_1 : UDINT := 16#0005_040C;    // 信息级槽 1（加减机延迟计时中） / info slot 1
    DL_CSM_CODE_INFO_2 : UDINT := 16#0005_040D;    // 信息级槽 2（供水低温保护强制减机） / info slot 2
    DL_CSM_CODE_FLT_1  : UDINT := 16#0005_0354;    // 故障级槽 1（无可用机组） / fault slot 1
    DL_CSM_CODE_FLT_2  : UDINT := 16#0005_0355;    // 故障级槽 2（负荷/台数组态非法） / fault slot 2
    DL_CSM_CODE_FLT_3  : UDINT := 16#0005_0356;    // 故障级槽 3（非有限/非法状态兜底） / fault slot 3
    DL_CSM_UNITS       : INT := 6;                 // 本件机组数，必须等于数组维度 [台] / Unit count, must match the arrays
    DL_CSM_DUTY_UNITS  : INT := 8;                 // 轮值件槽位数 [台] / Slot count of the duty block
    DL_CSM_DEMAND_MIN  : INT := 0;                 // 需求台数下限 [台] / Demand floor [pcs]
    DL_CSM_DEMAND_MAX  : INT := 6;                 // 需求台数上限 [台] / Demand ceiling [pcs]
    DL_CSM_IDX_NONE    : INT := -1;                // 无效机组号哨兵 [号] / Invalid unit sentinel
    DL_CSM_TAU_S       : LREAL := 60.0;            // 负荷率滤波时间常数 [s] / Load filter time constant [s]
    DL_CSM_PCT_MIN     : LREAL := 0.0;             // 百分数下限 [百分数] / Percent floor
    DL_CSM_PCT_MAX     : LREAL := 100.0;           // 百分数上限 [百分数] / Percent ceiling
    DL_CSM_DT_MIN_MS   : UDINT := 1;               // 扫描间隔下限 [ms]，防除零 / Scan interval floor [ms]
    DL_CSM_MS_PER_S    : LREAL := 1000.0;          // 毫秒转秒系数 [ms/s] / Milliseconds per second
    DL_CSM_ZERO        : LREAL := 0.0;             // 零值常量，避免裸字面量 [—] / Zero constant, avoids a bare literal
    DL_CSM_ONE         : LREAL := 1.0;             // 单位常量，滤波分子补项 [—] / Unity constant
    DL_CSM_TOL         : LREAL := 1.0E-6;          // 浮点比较容差 [—] / Float comparison tolerance
    DL_CSM_INF         : LREAL := 1.7976931348623157E308; // LREAL 幅值上限，Inf 判据 / LREAL magnitude ceiling
END_VAR

(*------------------------------------------------------------------------------
 * 段 1｜无条件刷新区（红线 5）：复位沿、两个延迟定时器与轮值件实例在任意分支之外
 *       周期调用恰好一次。轮值件按上一拍需求台数调度（单拍滞后对分钟级延迟无影响），
 *       保证使能/故障/各分支下轮值记账与最短时长保护永不断流
 *----------------------------------------------------------------------------*)
fbReset(CLK := bReset);                            // 复位沿检测无条件刷新 / reset edge refreshed unconditionally
fbTonUp(IN := bNeedUp AND (NOT bRearmUp), PT := tStageUpDelay);      // 加机延迟计时（重装拍强制复位）/ stage-up delay
fbTonDown(IN := bNeedDown AND (NOT bRearmDown), PT := tStageDownDelay);   // 减机延迟计时（重装拍强制复位）/ stage-down delay
IF bRearmUp THEN
    bRearmUp := FALSE;                             // 加机重装脉冲单拍自清 / re-arm pulse self-cleared
END_IF
IF bRearmDown THEN
    bRearmDown := FALSE;                           // 减机重装脉冲单拍自清 / re-arm pulse self-cleared
END_IF
FOR nLoop := 0 TO DL_CSM_DUTY_UNITS - 1 DO
    IF nLoop < DL_CSM_UNITS THEN
        abUnitReady[nLoop] := abChillerReady[nLoop];      // 0~5 槽接本件机组 / slots 0..5 map to the chillers
        abUnitRunning[nLoop] := abChillerRunning[nLoop];  // 运行反馈透传 / running feedback passed through
        abUnitFault[nLoop] := abChillerFault[nLoop];      // 故障透传（轮值件跳过）/ fault passed through
    ELSE
        abUnitReady[nLoop] := FALSE;               // 空槽：不就绪 / empty slot: not ready
        abUnitRunning[nLoop] := FALSE;             // 空槽：不运行 / empty slot: not running
        abUnitFault[nLoop] := FALSE;               // 空槽：不报故障（避免污染可用计数）/ empty slot: no fault
    END_IF
END_FOR
fbDuty(abUnitReady := abUnitReady,                 // 机组就绪（上限 8 槽）/ unit ready, 8 slots
       abUnitRunning := abUnitRunning,             // 运行反馈 / running feedback
       abUnitFault := abUnitFault,                 // 机组故障 / unit fault
       nDemand := nDemand,                         // 需求台数（上一拍生效值）[台] / demand of the previous scan
       bEnable := bEnable,                         // 使能透传 / enable forwarded
       uDeltaTimeMs := uDeltaTimeMs,               // 扫描间隔透传 [ms] / scan interval forwarded
       tMinRunTime := tMinRun,                     // 最小运行时长转发（时长逻辑归轮值件，不重复实现）/ min run forwarded
       tMinStopTime := tMinStop,                   // 最小停机时长转发 / min stop forwarded
       tRotateInterval := T#24H,                   // 轮值周期 24 小时（本件不另设引脚）/ rotation interval fixed at 24 h
       bForceRotate := FALSE,                      // 不强制轮值 / no forced rotation
       bReset := fbReset.Q,                        // 复位沿透传（R115：透传复位且只在故障相处置）/ reset edge forwarded
       abStartCmd => abStartCmdDuty,               // 轮值件启停命令暂存 / duty start commands staged
       nLeadUnit => nLeadStage,                    // 领机号暂存 / lead unit staged
       bError => bDutyFault);                      // 轮值件故障标志暂存（参数冲突透传）/ duty fault flag staged

(*------------------------------------------------------------------------------
 * 段 2｜复位沿处理（改写置于沿后，防吞沿 R39）：调度状态与需求台数回到保守初值
 *----------------------------------------------------------------------------*)
IF fbReset.Q THEN
    eState := E_DL_ChillerGroupState.eIdle;
    eErr   := 16#0000_0000;                        // 复位清码 / reset clears the code
    bError := FALSE;                               // 复位清故障 / reset clears the fault
    nDemand := DL_CSM_DEMAND_MIN;                  // 需求台数清 0 / demand cleared
    fLoadAvgPct := DL_CSM_ZERO;                    // 负荷率平滑值清 / smoothed load cleared
    bLowSupplyProtect := FALSE;                    // 低温保护标志清 / low-supply flag cleared
    bFirstScan := TRUE;                            // 重新首拍化 / re-initialize first scan
END_IF

(*------------------------------------------------------------------------------
 * 段 3｜机构闸（顺序判定，首个命中为准）：非有限 → 0356；组态非法 → 0355；
 *       无可用机组 → 0354。三者在同一个出口里全撤指令，避免多处 RETURN 漏赋值
 *----------------------------------------------------------------------------*)
bNonFin := (fSupplyC <> fSupplyC) OR (ABS(fSupplyC) >= DL_CSM_INF)
        OR (fReturnC <> fReturnC) OR (ABS(fReturnC) >= DL_CSM_INF)
        OR (fLoadPct <> fLoadPct) OR (ABS(fLoadPct) >= DL_CSM_INF)
        OR (fStageUpThrPct <> fStageUpThrPct) OR (ABS(fStageUpThrPct) >= DL_CSM_INF)
        OR (fStageDownThrPct <> fStageDownThrPct) OR (ABS(fStageDownThrPct) >= DL_CSM_INF)
        OR (fSupplyLowC <> fSupplyLowC) OR (ABS(fSupplyLowC) >= DL_CSM_INF);   // 引脚非有限汇总 / pins non-finite
nUsable := 0;                                      // 可用机组计数初值 / usable count seed
FOR nLoop := 0 TO DL_CSM_UNITS - 1 DO
    IF abChillerReady[nLoop] AND (NOT abChillerFault[nLoop]) THEN
        nUsable := nUsable + 1;                    // 就绪且无故障计入可用 [台] / usable unit counted
    END_IF
END_FOR
uGateCode := 16#0000_0000;                         // 机构闸码初值 0 / gate code seed
IF bNonFin THEN
    uGateCode := DL_CSM_CODE_FLT_3;                // 故障级：输入非有限（独立分支显式映射入 0356）/ fault: non-finite input
ELSIF (fStageDownThrPct >= fStageUpThrPct - DL_CSM_TOL)
   OR (fStageUpThrPct > DL_CSM_PCT_MAX + DL_CSM_TOL) OR (fStageUpThrPct < DL_CSM_PCT_MIN - DL_CSM_TOL)
   OR (fStageDownThrPct > DL_CSM_PCT_MAX + DL_CSM_TOL) OR (fStageDownThrPct < DL_CSM_PCT_MIN - DL_CSM_TOL) THEN
    uGateCode := DL_CSM_CODE_FLT_2;                // 故障级：阈值组态非法（减机阈值必须严格小于加机阈值）/ fault: threshold configuration invalid
ELSIF (nUsable < DL_CSM_DEMAND_MIN + 1) AND bEnable THEN
    uGateCode := DL_CSM_CODE_FLT_1;                // 故障级：无可用机组（工艺停机级）/ fault: no available unit, process stop level
END_IF
IF uGateCode <> 16#0000_0000 THEN
    eState := E_DL_ChillerGroupState.eFault;       // 进故障相 / enter fault state
    eErr   := uGateCode;                           // 落定机构闸码 / settle the gate code
    bError := TRUE;                                // 故障级必置 bError（R45 配对）/ fault-class pairs with bError
    bValid := FALSE;                               // 命令不可用 / commands unusable
    bNoAvailable := (uGateCode = DL_CSM_CODE_FLT_1);   // 无可用机组标志只在 0354 置位 / raised only on 0354
    bStageUpPending := FALSE;                      // 加机延迟标志撤 / stage-up pending withdrawn
    bStageDownPending := FALSE;                    // 减机延迟标志撤 / stage-down pending withdrawn
    FOR nLoop := 0 TO DL_CSM_UNITS - 1 DO
        abStartCmd[nLoop] := FALSE;                // 全撤启动命令安全侧 / every start command dropped
    END_FOR
    nRunningCmd := 0;                              // 指令台数清 / commanded count cleared
    nLeadChiller := DL_CSM_IDX_NONE;               // 领机号清 / lead cleared
    RETURN;
END_IF

(*------------------------------------------------------------------------------
 * 段 4｜负荷率一阶平滑：alpha = Δt / (tau + Δt)，时间常数 60 s。
 *       用注入间隔而非固定拍数，换任务周期不用改参数（跨平台可移植）
 *----------------------------------------------------------------------------*)
IF uDeltaTimeMs < DL_CSM_DT_MIN_MS THEN
    fDtSec := UDINT_TO_LREAL(DL_CSM_DT_MIN_MS) / DL_CSM_MS_PER_S;   // 间隔过小按下限 [s] / floored interval
ELSE
    fDtSec := UDINT_TO_LREAL(uDeltaTimeMs) / DL_CSM_MS_PER_S;       // 间隔原值 [s] / interval as-is
END_IF
fDenomSec := DL_CSM_TAU_S + fDtSec;                // 滤波分母 [s] / filter denominator [s]
IF fDenomSec > DL_CSM_TOL THEN
    fAlpha := fDtSec / fDenomSec;                  // 滤波系数（除子已判非零）[—] / filter coefficient
ELSE
    fAlpha := DL_CSM_ONE;                          // 分母异常：直通本拍值（不引入伪滤波）/ degenerate case passes through
END_IF
IF bFirstScan THEN
    fLoadAvgPct := fLoadPct;                       // 首拍直接取实测，避免从 0 爬升 / first scan takes the measurement
    bFirstScan := FALSE;                           // 首拍标志清除 / first-scan flag cleared
ELSE
    fLoadAvgPct := fLoadAvgPct + (fLoadPct - fLoadAvgPct) * fAlpha;   // 一阶平滑 [百分数] / first-order smoothing
END_IF

(*------------------------------------------------------------------------------
 * 段 5｜加/减机需求谓词与延迟（双延迟防抖动）：需求台数不超过可用台数；
 *       一次延迟周期只动一台，动作后强制重装定时器（负荷仍越限则再计一个周期）
 *----------------------------------------------------------------------------*)
bNeedUp := (fLoadAvgPct > fStageUpThrPct) AND (nDemand < nUsable);     // 加机需求：负荷高且还有可用机组 / stage-up need
bNeedDown := (fLoadAvgPct < fStageDownThrPct) AND (nDemand > DL_CSM_DEMAND_MIN);   // 减机需求：负荷低且还有机组在指令运行 / stage-down need
bStageUpPending := bNeedUp AND (NOT fbTonUp.Q);     // 加机延迟计时中 / stage-up delay running
bStageDownPending := bNeedDown AND (NOT fbTonDown.Q);   // 减机延迟计时中 / stage-down delay running
IF fbTonUp.Q THEN
    nDemand := nDemand + 1;                        // 加一台 [台] / stage up by one
    bRearmUp := TRUE;                              // 定时器重装，负荷仍高则再计一个周期 / re-arm for the next cycle
END_IF
IF fbTonDown.Q THEN
    nDemand := nDemand - 1;                        // 减一台 [台] / stage down by one
    bRearmDown := TRUE;                            // 定时器重装 / re-arm
END_IF

(*------------------------------------------------------------------------------
 * 段 6｜供水低温保护（防冻管）：低于门限强制再减一台，信息 040D。
 *       信息级不锁故障，但动作是强制的（安全侧：宁可欠冷，不可冻管）
 *----------------------------------------------------------------------------*)
bLowSupply := (fSupplyC < fSupplyLowC);            // 低温判据 [摄氏度] / low-supply predicate
bLowSupplyProtect := bLowSupply;                   // 保护标志出口 / protection flag outlet
IF bLowSupply AND (nDemand > DL_CSM_DEMAND_MIN) THEN
    nDemand := nDemand - 1;                        // 强制减一台 [台] / forced stage-down by one
END_IF

(*------------------------------------------------------------------------------
 * 段 7｜需求台数域钳位（0~6 且不超可用台数）：域外一律钳，不新占码位
 *----------------------------------------------------------------------------*)
IF nDemand < DL_CSM_DEMAND_MIN THEN
    nDemand := DL_CSM_DEMAND_MIN;                  // 下限钳位 / clipped to the floor
END_IF
IF nDemand > DL_CSM_DEMAND_MAX THEN
    nDemand := DL_CSM_DEMAND_MAX;                  // 上限钳位 / clipped to the ceiling
END_IF
IF nDemand > nUsable THEN
    nDemand := nUsable;                            // 不超过可用台数（故障切备后的自然收敛）/ clamped to the usable count
END_IF
IF bEnable AND (nDemand < DL_CSM_DEMAND_MIN + 1) THEN
    nDemand := DL_CSM_DEMAND_MIN + 1;              // 使能保底一台领机（否则 10 分钟无冷才起动，工艺不可接受）/ at least one chiller when enabled
END_IF

(*------------------------------------------------------------------------------
 * 段 8｜轮值件故障透传（R115）：只在故障相处置，下一步由 CASE 的 eFault 分支承接
 *----------------------------------------------------------------------------*)
IF bDutyFault THEN
    eState := E_DL_ChillerGroupState.eFault;       // 轮值件参数冲突：进故障相 / duty parameter conflict enters fault
    eErr   := DL_CSM_CODE_FLT_2;                   // 复用组态非法槽（台数/参数冲突同一出口，不升格不加码）/ reuses the configuration slot
    bError := TRUE;                                // 故障级必置 bError（R45 配对）/ fault-class pairs with bError
    bValid := FALSE;                               // 命令不可用 / commands unusable
END_IF

(*------------------------------------------------------------------------------
 * 段 9｜状态机：CASE 含 ELSE 兜底（非法状态 → 0356 + 全撤指令）
 *----------------------------------------------------------------------------*)
CASE eState OF

    E_DL_ChillerGroupState.eIdle:
        bValid := FALSE;                           // 失能闸显式不可用（R72）/ explicit FALSE on the disable gate
        bNoAvailable := FALSE;                     // 无可用标志撤 / no-available flag withdrawn
        bLowSupplyProtect := FALSE;                // 低温保护标志撤 / low-supply flag withdrawn
        bStageUpPending := FALSE;                  // 加机延迟标志撤 / stage-up pending withdrawn
        bStageDownPending := FALSE;                // 减机延迟标志撤 / stage-down pending withdrawn
        eErr := 16#0000_0000;                      // 待机无错 / no error in idle
        bError := FALSE;                           // 待机无故障 / no fault in idle
        IF bEnable THEN
            eState := E_DL_ChillerGroupState.eRunning;   // 使能进稳态调度 / enable enters steady scheduling
        END_IF

    E_DL_ChillerGroupState.eRunning:
        bValid := TRUE;                            // 命令可用 / commands usable
        bError := FALSE;                           // 稳态无故障 / no fault in the steady state
        eErr := 16#0000_0000;                      // 稳态先清码 / clear the code first
        IF bLowSupplyProtect THEN
            eErr := DL_CSM_CODE_INFO_2;            // 信息级：供水低温保护强制减机（优先）/ info: low-supply protection outranks the delay hint
            eState := E_DL_ChillerGroupState.eLowSupply;   // 转低温保护相 / enter the protection state
        ELSIF bStageUpPending THEN
            eErr := DL_CSM_CODE_INFO_1;            // 信息级：加机延迟计时中 / info: stage-up delay running
            eState := E_DL_ChillerGroupState.eStageUp;     // 转加机延迟相 / enter the stage-up state
        ELSIF bStageDownPending THEN
            eErr := DL_CSM_CODE_INFO_1;            // 信息级：减机延迟计时中 / info: stage-down delay running
            eState := E_DL_ChillerGroupState.eStageDown;   // 转减机延迟相 / enter the stage-down state
        END_IF
        IF NOT bEnable THEN
            eState := E_DL_ChillerGroupState.eIdle;    // 失能回待机 / disable returns to idle
            bValid := FALSE;                       // 失能闸显式不可用 / explicit FALSE on the disable gate
        END_IF

    E_DL_ChillerGroupState.eStageUp:
        bValid := TRUE;                            // 命令可用（延迟期内照常调度）/ commands usable during the delay
        bError := FALSE;                           // 信息级不置 bError / info never raises bError
        eErr := DL_CSM_CODE_INFO_1;                // 信息级：加机延迟计时中 / info: stage-up delay running
        IF NOT bEnable THEN
            eState := E_DL_ChillerGroupState.eIdle;    // 失能回待机（退出条件一）/ disable, first exit
            bValid := FALSE;                       // 失能闸显式不可用 / explicit FALSE on the disable gate
        ELSIF bLowSupplyProtect THEN
            eState := E_DL_ChillerGroupState.eLowSupply;   // 低温保护优先（退出条件二）/ protection outranks, second exit
        ELSIF (NOT bNeedUp) THEN
            eState := E_DL_ChillerGroupState.eRunning;     // 负荷回落回稳态（退出条件三）/ load fell back, third exit
        END_IF

    E_DL_ChillerGroupState.eStageDown:
        bValid := TRUE;                            // 命令可用 / commands usable
        bError := FALSE;                           // 信息级不置 bError / info never raises bError
        eErr := DL_CSM_CODE_INFO_1;                // 信息级：减机延迟计时中 / info: stage-down delay running
        IF NOT bEnable THEN
            eState := E_DL_ChillerGroupState.eIdle;    // 失能回待机（退出条件一）/ disable, first exit
            bValid := FALSE;                       // 失能闸显式不可用 / explicit FALSE on the disable gate
        ELSIF bLowSupplyProtect THEN
            eState := E_DL_ChillerGroupState.eLowSupply;   // 低温保护优先（退出条件二）/ protection outranks, second exit
        ELSIF (NOT bNeedDown) THEN
            eState := E_DL_ChillerGroupState.eRunning;     // 负荷回升回稳态（退出条件三）/ load recovered, third exit
        END_IF

    E_DL_ChillerGroupState.eLowSupply:
        bValid := TRUE;                            // 命令可用（保护动作已强制减机）/ commands usable after the forced stage-down
        bError := FALSE;                           // 信息级不锁故障 / info never latches a fault
        eErr := DL_CSM_CODE_INFO_2;                // 信息级：供水低温保护强制减机 / info: forced stage-down on low supply
        IF NOT bEnable THEN
            eState := E_DL_ChillerGroupState.eIdle;    // 失能回待机（退出条件一）/ disable, first exit
            bValid := FALSE;                       // 失能闸显式不可用 / explicit FALSE on the disable gate
        ELSIF (NOT bLowSupplyProtect) THEN
            eState := E_DL_ChillerGroupState.eRunning; // 供水温度回升回稳态（退出条件二）/ supply recovered, second exit
        END_IF

    E_DL_ChillerGroupState.eFault:
        bValid := FALSE;                           // 故障闸显式不可用（R72）/ explicit FALSE on the fault gate
        bError := TRUE;                            // 故障级必置 bError（R45 配对）/ fault-class pairs with bError
        bStageUpPending := FALSE;                  // 加机延迟标志撤 / stage-up pending withdrawn
        bStageDownPending := FALSE;                // 减机延迟标志撤 / stage-down pending withdrawn
        IF eErr = 16#0000_0000 THEN
            eErr := DL_CSM_CODE_FLT_3;             // 入口无码时按非法状态兜底（R45：bError 必须有对应码）/ illegal-state fallback
        END_IF
        IF bEnable AND (NOT bDutyFault) AND (nUsable >= DL_CSM_DEMAND_MIN + 1)
           AND (fStageDownThrPct < fStageUpThrPct - DL_CSM_TOL) THEN
            eState := E_DL_ChillerGroupState.eIdle;    // 前置条件全部恢复才回待机（退出条件 ≥2）/ recover only when every precondition is back
        END_IF

    ELSE
        eState := E_DL_ChillerGroupState.eFault;    // 非法状态兜底 / illegal-state fallback
        eErr := DL_CSM_CODE_FLT_3;                 // 故障级兜底：非法状态 / fault fallback: illegal state
        bError := TRUE;                            // 故障级必置 bError（R45 配对）/ fault-class pairs with bError
        bValid := FALSE;                           // 命令不可用 / commands unusable
        bStageUpPending := FALSE;                  // 加机延迟标志撤 / stage-up pending withdrawn
        bStageDownPending := FALSE;                // 减机延迟标志撤 / stage-down pending withdrawn

END_CASE

(*------------------------------------------------------------------------------
 * 段 10｜出口装配：轮值件命令落到 0~5 号池、领机号映射、指令台数统计；
 *        失能/故障一律全撤（安全值而非上次值，红线 6）
 *----------------------------------------------------------------------------*)
nRunningCmd := 0;                                  // 指令台数从零重数 / commanded count recounted
FOR nLoop := 0 TO DL_CSM_UNITS - 1 DO
    IF bEnable AND bValid THEN
        abStartCmd[nLoop] := abStartCmdDuty[nLoop];     // 正常调度：透传轮值件命令 / pass the duty command through
    ELSE
        abStartCmd[nLoop] := FALSE;                     // 失能/故障：全撤安全侧 / drop everything, safe side
    END_IF
    IF abStartCmd[nLoop] THEN
        nRunningCmd := nRunningCmd + 1;                 // 指令台数累加 [台] / commanded count increments
    END_IF
END_FOR
IF (nLeadStage >= 0) AND (nLeadStage < DL_CSM_UNITS) AND bEnable AND bValid THEN
    nLeadChiller := nLeadStage;                    // 领机号映射（空槽不冒充）/ lead mapped, empty slots never pose as a lead
ELSE
    nLeadChiller := DL_CSM_IDX_NONE;               // 无领机 / no lead chiller
END_IF
END_FUNCTION_BLOCK

(* ---- FB_DL_ChillerStagingCurve.st ---- *)
(*==============================================================================
 * 组件名称 (Component)  : FB_DL_ChillerStagingCurve
 * 所属子库 (Sublibrary) : DL_Process
 * 当前版本 (Version)    : 1.0.1
 * 兼容性 (Platform)     : CODESYS 3.5 / TwinCAT 3 / 汇川 InoProShop（纯标准元素，无方言）
 * 功能描述 (Function)   : 冷机加减机效率曲线选点。用单机 COP 与容量曲线求最经济负荷点，
 *                         按系统负荷率反算建议台数（N+1 冗余口径：需求台数向上取整再加一台，
 *                         下限钳 1 台、上限 8 台），与在线台数比较后在死区外、持续确认时长
 *                         满足时给单拍加/减机请求。曲线非单调或含非有限值一律**不给建议**
 *                         （错曲线的建议比不给更危险）。不做机组启停时序、不做 COP 实测、
 *                         不做负荷预测。
 *                         交付门槛：本件不含时间转换链，纯实数与整数算术，无平台相关内建。
 * 溯源 (Origin)         : 道莅 clean-room 防御性实现
 * 本文件内含 (Contains) : TYPE E_DL_StageState / FUNCTION_BLOCK FB_DL_ChillerStagingCurve
 * 依赖 (Depends)        : 无（仅 Standard.library 的 ABS / LIMIT / TRUNC）
 * 红线自检 (Redline)    : 无外部全局变量、无硬件地址直引 ｜ 全变量中英双语同行注释
 *                         台数判零防除零 ｜ 曲线单调性与非有限双检 ｜ 负荷非有限保持上次台数 ｜
 *                         确认定时器与沿实例无条件周期刷新 ｜ 枚举显式赋值 ｜ CASE 含 ELSE
 * 错误码表 (Codes)      : 16#0005_0449 就绪（建议已给出且曲线有效）
 *                         16#0005_044A 预留：本版不发码（下一轮区间起点，禁止回填）
 *                         16#0005_044B 故障级 曲线非单调或含非有限值，不给建议
 *                         16#0005_044C 故障级 在线台数为 0（防除零，不给建议）
 *                         16#0005_044D 信息级 负荷率非有限，保持上次台数与 COP（不置故障级标志）
 * 修订历史 (Revision)   : 2026-11-17  v1.0.0  首版入库 · R28 · 阶段三批 4
 *                         2026-11-17  v1.0.1  终审修复：①需求台数向上取整算式在「正好整除」
 *                                    时多算一台（TRUNC+1 把整数也进位了），改为余量判进位；
 *                                    ②负荷率与死区补域钳制（超界负荷经实数转整数溢出会让加减
 *                                    机方向翻转）；③故障解除判据原写成「失能且未锁存」永不成立，
 *                                    改为失能即解除（原写法使组态类故障永久不可恢复）· R28 · 阶段四
 * 验收向量 (Acceptance) : 正向 负荷 55 %、在线 3 台、曲线峰值在 80 %（单机 18.3 % 过轻）→
 *                         bDelReq 单拍、uStage=2、bOnCurve=TRUE
 *                         反向 曲线改为非单调 → 16#0005_044B 且 bAddReq/bDelReq 均为 FALSE；
 *                         台数给 0 → 16#0005_044C；负荷给 NaN → 16#0005_044D 且 uStage 保持
 *============================================================================*)

(*-----------------------------------------------------------------------------
 * 枚举: E_DL_StageState（归属本功能块，同文件发布，全库唯一定义）
 *----------------------------------------------------------------------------*)
TYPE E_DL_StageState :
(
    eIdle    := 0,    // 待机：使能关或曲线无效 / Idle, disabled or the curve is invalid
    eEval    := 10,   // 评估：本拍算建议台数 / Evaluating the recommended unit count
    eConfirm := 20,   // 确认：偏差持续计时中 / Confirming, the deviation persists
    ePulse   := 30,   // 脉冲：本拍发出加/减机请求 / Pulse, an add or delete request is issued this scan
    eFault   := 99    // 故障：锁存码保持 / Fault, the latch code is held
);
END_TYPE

FUNCTION_BLOCK FB_DL_ChillerStagingCurve
VAR_INPUT
    bEnable       : BOOL := FALSE;        // 使能 / Enable
    fLoadPct      : REAL := 50.0;         // 系统负荷率 [%]，域 0~120 / System load in percent, domain 0 to 120
    afCopCurve    : ARRAY[1..11] OF REAL; // 单机 COP 曲线（10/20/…/100 % 十一点） / Single-unit COP curve, eleven points
    afCapCurve    : ARRAY[1..11] OF REAL; // 单机容量曲线 [kW]（十一点） / Single-unit capacity curve in kilowatt
    uUnitCnt      : UINT := 2;            // 在线台数 [台]，域 1~8 / Online unit count, domain 1 to 8
    fLoadStepPct  : REAL := 5.0;          // 加/减机死区 [%]，域 1~20 / Staging dead band in percent, domain 1 to 20
    tConfirm      : TIME := T#60S;        // 建议持续确认 [ms]，域 10 s~10 min / Suggestion confirmation time
END_VAR
VAR_OUTPUT
    uStage        : UINT := 1;            // 建议运行台数 [台]，域 1~8 / Recommended unit count
    bAddReq       : BOOL;                 // 加机请求（单拍脉冲） / Add request, a one-scan pulse
    bDelReq       : BOOL;                 // 减机请求（单拍脉冲） / Delete request, a one-scan pulse
    fCopNow       : REAL;                 // 当前负荷率推算 COP / COP derived from the present per-unit load
    fBestLoadPct  : REAL;                 // 本台数最经济负荷率 [%] / Most economic per-unit load
    bOnCurve      : BOOL;                 // 曲线单调性校验通过 / Curve monotonicity check passed
    eErr          : UDINT;                // 错误码，段位 16#0005_xxxx / Error code in segment 16#0005_xxxx
END_VAR
VAR
    _eState       : E_DL_StageState := E_DL_StageState.eIdle; // 当前相位 / Current phase
    _bInit        : BOOL := FALSE;        // 首扫标志，取非判定 / First-scan flag, tested negated
    _bCurveOk     : BOOL;                 // 曲线有效标志 / Curve valid flag
    _bLoadOk      : BOOL;                 // 负荷有限标志 / Load finite flag
    _bUpWant      : BOOL;                 // 需要加机（未确认） / Add needed before confirmation
    _bDnWant      : BOOL;                 // 需要减机（未确认） / Delete needed before confirmation
    _bFaultLatch  : BOOL := FALSE;        // 故障锁存标志 / Fault latch flag
    _uLatchCode   : UDINT;                // 锁存码载体 / Latch code carrier
    _uStageCalc   : UINT := 1;            // 本拍计算建议台数 [台] / Computed recommended count
    _uBestIdx     : UINT := 11;           // COP 峰值点下标（10..100 %） / Index of the COP peak
    _uStagePrev   : UINT := 1;            // 上次台数（非有限负荷时保持） / Previous count kept for a non-finite load
    _iLoop        : INT;                  // 曲线扫描索引 / Curve scan index
    _iGuard       : INT;                  // 防死循环计数器 / Loop guard counter
    _fBestCop     : REAL := 0.0;          // 峰值 COP / Peak COP
    _fPerUnit     : REAL;                 // 单机负荷率 [%] / Per-unit load in percent
    _fLoadEff     : REAL;                 // 域钳制后负荷率 [%]（0~120） / Load after the domain clamp
    _fStepEff     : REAL := 5.0;          // 域钳制后死区 [%]（1~20） / Dead band after the domain clamp
    _fNeedUnits   : REAL;                 // 需求台数（未取整） / Required unit count before rounding
    _fCopLocal    : REAL;                 // 当前 COP 插值结果 / Interpolated COP
    _rtrigConf    : R_TRIG;               // 确认计时满上升沿 / Rising edge of the confirmation timer
    _tonConfirm   : TON;                  // 建议持续确认计时 / Suggestion confirmation timer
END_VAR
VAR CONSTANT
    DL_CH_READY    : UDINT := 16#0005_0449;  // 就绪码 / Ready code
    DL_CH_CURVE_BAD : UDINT := 16#0005_044B; // 故障级曲线不可用码 / Fault code for an unusable curve
    DL_CH_UNIT_ZERO : UDINT := 16#0005_044C; // 故障级台数为零码 / Fault code for a zero unit count
    DL_CH_LOAD_BAD : UDINT := 16#0005_044D;  // 信息级负荷非有限码 / Info code for a non-finite load
    DL_CH_PTS      : INT := 11;              // 曲线点数 / Curve point count
    DL_CH_LOOP_MAX : INT := 20;              // 循环保护上限 / Loop guard bound
    DL_CH_STEP_LO  : REAL := 1.0;            // 死区下限 [%] / Dead band lower bound
    DL_CH_STEP_HI  : REAL := 20.0;           // 死区上限 [%] / Dead band upper bound
    DL_CH_STEP_DFLT : REAL := 5.0;           // 死区非有限时的默认值 [%] / Default dead band for a non-finite input
    DL_CH_LOAD_HI  : REAL := 120.0;          // 负荷率域上限 [%] / Load domain upper bound
    DL_CH_NEED_HI  : REAL := 100.0;          // 需求台数兜底上限 [台] / Required-unit upper bound guard
    DL_CH_STAGE_LO : UINT := 1;              // 建议台数下限 [台] / Recommended count lower bound
    DL_CH_STAGE_HI : UINT := 8;              // 建议台数上限 [台] / Recommended count upper bound
    DL_CH_UNIT_MAX : UINT := 8;              // 在线台数上限 [台] / Online count upper bound
    DL_CH_EPS      : REAL := 1.0E-6;         // 浮点判零容差 / Float zero tolerance
END_VAR

// 段 1｜输出与单拍标志预置
bAddReq := FALSE;                                   // 加机请求预清（单拍） / Add request pre-cleared
bDelReq := FALSE;                                   // 减机请求预清（单拍） / Delete request pre-cleared
bOnCurve := FALSE;                                  // 曲线校验标志预清 / Curve check flag pre-cleared
eErr := 0;                                          // 错误码预清 / Error code pre-cleared
_fCopLocal := 0.0;                                  // COP 局部量预清 / COP local pre-cleared

// 段 2｜确认定时器与沿实例无条件周期刷新
_tonConfirm(IN := bEnable AND _bCurveOk AND (_bUpWant OR _bDnWant), PT := tConfirm);
_rtrigConf(CLK := _tonConfirm.Q);                   // 确认满沿 / Confirmation edge

// 段 3｜首扫初始化（判据取非，R19）
IF NOT _bInit THEN
    uStage := 1;                                    // 建议台数起点 1 [台] / Recommended count starts at one
    _uStagePrev := 1;
    _eState := E_DL_StageState.eIdle;               // 相位待机起步 / Phase starts idle
    _bInit := TRUE;                                 // 首扫只做一次 / The first scan runs once
END_IF

// 段 4｜曲线校验（单调不减 + 全点有限；十一轮固定上界，循环带保护计数）
_bCurveOk := TRUE;
_iLoop := 1;
_iGuard := 0;
_fBestCop := 0.0 - 1.0E30;
_uBestIdx := 1;
WHILE (_iLoop <= DL_CH_PTS) AND (_iGuard < DL_CH_LOOP_MAX) DO
    IF (afCopCurve[_iLoop] <> afCopCurve[_iLoop]) OR ((afCopCurve[_iLoop] - afCopCurve[_iLoop]) <> (afCopCurve[_iLoop] - afCopCurve[_iLoop])) THEN
        _bCurveOk := FALSE;                         // COP 点非有限 / A COP point is not finite
    END_IF
    IF (afCapCurve[_iLoop] <> afCapCurve[_iLoop]) OR ((afCapCurve[_iLoop] - afCapCurve[_iLoop]) <> (afCapCurve[_iLoop] - afCapCurve[_iLoop])) THEN
        _bCurveOk := FALSE;                         // 容量点非有限 / A capacity point is not finite
    END_IF
    IF afCopCurve[_iLoop] > _fBestCop THEN
        _fBestCop := afCopCurve[_iLoop];            // 峰值刷新 / Peak refreshed
        _uBestIdx := INT_TO_UINT(_iLoop);           // 峰值下标 / Peak index
    END_IF
    IF _iLoop > 1 THEN
        IF afCopCurve[_iLoop] < afCopCurve[_iLoop - 1] THEN
            _bCurveOk := FALSE;                     // 非单调（COP 随负荷率不增）：不给建议 / Non-monotonic curve, no advice
        END_IF
        IF afCapCurve[_iLoop] < afCapCurve[_iLoop - 1] THEN
            _bCurveOk := FALSE;                     // 容量曲线非单调 / Non-monotonic capacity curve
        END_IF
    END_IF
    _iLoop := _iLoop + 1;
    _iGuard := _iGuard + 1;                         // 防死循环计数 / Loop guard incremented
END_WHILE
bOnCurve := _bCurveOk;                              // 曲线校验出口 / Curve check output
fBestLoadPct := UINT_TO_REAL(_uBestIdx) * 10.0;     // 最经济负荷率 [%] / Most economic load
IF NOT _bCurveOk THEN
    eErr := DL_CH_CURVE_BAD;                        // 故障级：曲线不可用 / Fault, the curve is unusable
    _uLatchCode := DL_CH_CURVE_BAD;
    _bFaultLatch := TRUE;
    _eState := E_DL_StageState.eFault;
END_IF

// 段 5｜台数与负荷闸（台数 0 防除零；负荷非有限保持上次台数）
IF uUnitCnt = 0 THEN
    eErr := DL_CH_UNIT_ZERO;                        // 故障级：在线台数为 0 / Fault, the online unit count is zero
    _uLatchCode := DL_CH_UNIT_ZERO;
    _bFaultLatch := TRUE;
    _eState := E_DL_StageState.eFault;
END_IF
_bLoadOk := NOT ((fLoadPct <> fLoadPct) OR ((fLoadPct - fLoadPct) <> (fLoadPct - fLoadPct)));
IF NOT _bLoadOk THEN
    eErr := DL_CH_LOAD_BAD;                         // 信息级：负荷非有限，保持上次台数 / Info, the load is not finite and the previous count is held
    uStage := _uStagePrev;
END_IF

// 段 6｜建议台数计算（N+1 冗余口径：需求台数向上取整再加 1 台，钳 1~8）
IF _bCurveOk AND _bLoadOk AND (uUnitCnt > 0) AND (fBestLoadPct > DL_CH_EPS) THEN
    _fLoadEff := LIMIT(0.0, fLoadPct, DL_CH_LOAD_HI);   // 负荷率域钳制 [%]（防实数转整数溢出翻转加减机方向） / Load clamped into the domain
    _fStepEff := fLoadStepPct;                          // 死区副本 [%] / Dead band copy
    IF (_fStepEff <> _fStepEff) OR ((_fStepEff - _fStepEff) <> (_fStepEff - _fStepEff)) THEN
        _fStepEff := DL_CH_STEP_DFLT;                   // 死区非有限：回默认值，不静默变成 0 死区 / Non-finite dead band falls back to the default
    END_IF
    _fStepEff := LIMIT(DL_CH_STEP_LO, _fStepEff, DL_CH_STEP_HI);   // 死区域钳制 [%] / Dead band clamped
    _fPerUnit := _fLoadEff / UINT_TO_REAL(uUnitCnt);    // 单机负荷率 [%] / Per-unit load
    _fNeedUnits := _fLoadEff / fBestLoadPct;            // 需求台数（未取整） / Required units before rounding
    IF _fNeedUnits < 0.0 THEN
        _fNeedUnits := 0.0;                             // 负负荷按 0 处理 / Negative load treated as zero
    END_IF
    IF _fNeedUnits > DL_CH_NEED_HI THEN
        _fNeedUnits := DL_CH_NEED_HI;                   // 上限兜底，防取整溢出 [台] / Upper bound guard against rounding overflow
    END_IF
    _uStageCalc := REAL_TO_UINT(TRUNC(_fNeedUnits));    // 先向下取整 [台] / Truncate first
    IF _fNeedUnits > UINT_TO_REAL(_uStageCalc) THEN
        _uStageCalc := _uStageCalc + 1;                 // 有小数余量才进一位（正好整除不进位） / Round up only with a fractional remainder
    END_IF
    _uStageCalc := _uStageCalc + 1;                     // N+1 冗余 [台] / One redundant unit
    uStage := LIMIT(DL_CH_STAGE_LO, _uStageCalc, DL_CH_STAGE_HI); // 建议台数钳制 [台] / Recommended count clamped
    _uStagePrev := uStage;                          // 台数快照 / Count snapshot
    // 当前负荷率下的 COP 插值（十一点等距，线性内插）
    IF _fPerUnit <= 10.0 THEN
        _fCopLocal := afCopCurve[1];                // 低于首点：取首点 / Below the first point, use the first
    ELSIF _fPerUnit >= 100.0 THEN
        _fCopLocal := afCopCurve[11];               // 高于末点：取末点 / Above the last point, use the last
    ELSE
        _iLoop := TRUNC(_fPerUnit / 10.0) + 1;      // 区间左端下标 / Left index of the interval
        IF _iLoop < 1 THEN
            _iLoop := 1;                            // 下标下限保护 / Index lower guard
        END_IF
        IF _iLoop > (DL_CH_PTS - 1) THEN
            _iLoop := DL_CH_PTS - 1;                // 下标上限保护 / Index upper guard
        END_IF
        _fCopLocal := afCopCurve[_iLoop]
                    + ((afCopCurve[_iLoop + 1] - afCopCurve[_iLoop])
                       * ((_fPerUnit - (UINT_TO_REAL(INT_TO_UINT(_iLoop)) * 10.0) + 10.0) / 10.0 - 1.0));
    END_IF
    fCopNow := _fCopLocal;                          // COP 出口 / COP output
    // 死区比较：死区外才提请求（防抖）
    _bUpWant := (_fPerUnit > (fBestLoadPct + _fStepEff)) OR (uStage > uUnitCnt);
    _bDnWant := ((_fPerUnit < (fBestLoadPct - _fStepEff)) OR (uStage < uUnitCnt)) AND (uStage >= DL_CH_STAGE_LO);
    IF uStage > uUnitCnt THEN
        _bUpWant := TRUE;                           // 建议台数高于在线台数：加机 / The recommendation exceeds the online count
        _bDnWant := FALSE;
    ELSIF uStage < uUnitCnt THEN
        _bUpWant := FALSE;                          // 建议台数低于在线台数：减机 / The recommendation is below the online count
        _bDnWant := TRUE;
    ELSE
        _bUpWant := FALSE;                          // 台数一致：不提请求 / Counts agree, no request
        _bDnWant := FALSE;
    END_IF
    eErr := DL_CH_READY;                            // 就绪码 / Ready code
END_IF

// 段 7｜请求脉冲（确认时长满才发，单拍自清）
IF (_eState <> E_DL_StageState.eFault) THEN
    IF _rtrigConf.Q THEN
        IF _bUpWant AND (uUnitCnt < DL_CH_UNIT_MAX) THEN
            bAddReq := TRUE;                        // 加机单拍脉冲 / Add pulse for one scan
        ELSIF _bDnWant AND (uUnitCnt > DL_CH_STAGE_LO) THEN
            bDelReq := TRUE;                        // 减机单拍脉冲（下限钳 1 台） / Delete pulse, the count is clamped to one
        END_IF
        _eState := E_DL_StageState.ePulse;          // 本拍脉冲相 / Pulse phase for this scan
    ELSE
        IF bEnable AND _bCurveOk AND _bLoadOk THEN
            IF _bUpWant OR _bDnWant THEN
                _eState := E_DL_StageState.eConfirm;    // 偏差存在：确认计时中 / Deviation present, confirming
            ELSE
                _eState := E_DL_StageState.eEval;       // 无偏差：常规评估 / No deviation, plain evaluation
            END_IF
        ELSE
            _eState := E_DL_StageState.eIdle;           // 禁用或输入不可用：待机 / Disabled or unusable inputs, idle
        END_IF
    END_IF
END_IF

// 段 8｜相位收口（ENUM + CASE + ELSE 兜底）
CASE _eState OF
    E_DL_StageState.eIdle:
        bAddReq := FALSE;                           // 待机不发请求 / No request while idle
        bDelReq := FALSE;
    E_DL_StageState.eEval:
        bAddReq := FALSE;                           // 评估相不发请求 / No request while evaluating
        bDelReq := FALSE;
    E_DL_StageState.eConfirm:
        bAddReq := FALSE;                           // 确认相不发请求 / No request while confirming
        bDelReq := FALSE;
    E_DL_StageState.ePulse:
        _eState := E_DL_StageState.eEval;           // 脉冲相单拍后自动转评估 / The pulse phase lasts one scan
    E_DL_StageState.eFault:
        bAddReq := FALSE;                           // 故障相不发请求 / No request in the fault phase
        bDelReq := FALSE;
        eErr := _uLatchCode;                        // 锁存码回放 / Replay the latch code
        IF NOT bEnable THEN                         // 失能即解除锁存（旧判据取反写错，故障永不可退） / A disable releases the latch
            _bFaultLatch := FALSE;                  // 锁存解除 / Latch released
            _uLatchCode := 0;                       // 锁存码清 / Latch code cleared
            eErr := DL_CH_READY;                    // 解除后回就绪码 / Ready code after the release
            _eState := E_DL_StageState.eIdle;       // 回待机 / Back to idle
        END_IF
    ELSE
        // 非法相位兜底（故障级）
        bAddReq := FALSE;
        bDelReq := FALSE;
        eErr := DL_CH_CURVE_BAD;                    // 故障级：非法相位 / Fault, illegal phase
        _uLatchCode := DL_CH_CURVE_BAD;
        _bFaultLatch := TRUE;
        _eState := E_DL_StageState.eFault;
END_CASE
END_FUNCTION_BLOCK

(* ---- FB_DL_ChillerStagingSeq.st ---- *)
(*
  组件名 Component   : FB_DL_ChillerStagingSeq
  子库 Sublibrary    : DL_Process
  版本 Version       : 1.0.0
  兼容性 Platform    : CODESYS 3.5 / TwinCAT 3 / 汇川 InoProShop / Machine Expert（仅 Standard.library）
  功能 Function      : 冷机加卸载顺控（与 ChillerTempStab/ChillerCondReset 分工：稳定
                       判稳 vs 顺控编组）：
                       1) 按需量 nDemand 分级加/卸载：在编台数 < 需量 → 启动累计运行
                       时间最短的停机台；> 需量 → 停止累计运行时间最长的运行台（轮值
                       均衡按运行小时数自然轮换）；
                       2) 最短启停驻留：每台独立启停驻留扫描计数，未满驻留不得启停，
                       驻留阻塞期置 bDwellLock（信息级）；
                       3) 需量越域钳位 [0, 台数上限] 并留信息码（瞬时口径）；
                       4) 到期轮值检查窗自复触周期计时（R188 范式）。
  边界 Boundary      : ① 本件只出各台启停指令，不写物理 IO，不接管冷冻水回路；
                       ② 运行时间累计由本件按扫描期内部折算（tCycle 换算分钟），
                       上位机无需另喂运行时数；
                       ③ 故障锁存解除唯一路径 = bReset 上升沿（输入引脚，恒可达）；
                       ④ 无全局变量引用、无外部变量声明、无物理地址寻址。
  依赖 Depends       : Standard.library（R_TRIG / TON）
  溯源 Origin        : 道莅自研 clean-room（参考 t2-7-packml 最小子集与 t1-2-oscat
                       暖通语义分类与参数域，零代码行复制）
  码位 Code          : 16#06_0_BD（Process 段 0006，B 子带 BD 格）
  码表 Error codes（本件格 06_0_BD，单轨子道：故障 0x02BD / 信息 0x01BD）:
    16#0006_02BD 故障级：组态非法（台数越域 / 驻留或周期为 0），锁存至复位
    16#0006_01BD 信息级：需量越域已钳位（瞬时口径，不置 bError）
  修订历史 Revision  :
    2026-11-19  v1.0.0  R44 首版（批次 3 · 序号 14）
*)

TYPE E_DL_CssState :
(
    eIdle  := 0,    // 空闲：未使能，全台停机 / Idle, all stages off
    eRun   := 10,   // 编组运行：加卸载顺控 / Running, staging sequence
    eFault := 90    // 故障：组态锁存 / Fault, latched
);
END_TYPE

FUNCTION_BLOCK FB_DL_ChillerStagingSeq
VAR_INPUT
    bEnable  : BOOL;                       // 使能（电平）[-] / Enable
    bReset   : BOOL;                       // 上升沿清故障锁存 [-] / Reset edge
    nDemand  : INT;                        // 需量台数 [台]，域 0..4 / Required stage count
    tMinOn   : TIME := T#300S;             // 最短运行驻留 [毫秒] / Minimum on dwell
    tMinOff  : TIME := T#600S;             // 最短停机驻留 [毫秒] / Minimum off dwell
    tRotateWin: TIME := T#60S;             // 轮值均衡检查窗 [毫秒] / Rotation check window
    tCycle   : TIME := T#1S;               // 扫描周期 [毫秒] / Scan cycle time
END_VAR
VAR_OUTPUT
    abStageRun : ARRAY[1..4] OF BOOL;      // 各台运行指令输出 [-] / Stage run commands
    nStaged    : INT;                      // 在编台数 [台] / Staged count
    bDwellLock : BOOL;                     // 驻留阻塞电平 [-] / Dwell blocking level
    eState     : E_DL_CssState;            // 状态出口，段尾单点映射 / State outlet
    bError     : BOOL;                     // 故障锁存标志 [-] / Fault latch flag
    uErrId     : UDINT;                    // 事件码，0 = 无事件 / Event code
END_VAR
VAR
    rtReset : R_TRIG;                      // 复位沿实例，段 0 无条件刷新 / Reset edge
    tonRotateWin: TON;                     // 轮值检查窗（自复触，R188） / Rotation window
    _eState : E_DL_CssState := E_DL_CssState.eIdle;    // 内部相位（CASE 唯一写入目标）/ Internal phase
    _nDemandUse: INT;                      // 钳位后需量 [台] / Clamped demand
    _auRunMin  : ARRAY[1..4] OF UDINT;     // 各台累计运行时间 [分] / Runtime per stage
    _auDwellScan: ARRAY[1..4] OF UDINT;    // 各台启停驻留扫描计 [拍] / Dwell scans per stage
    _abLastRun : ARRAY[1..4] OF BOOL;      // 各台上拍运行态镜像 [-] / Previous run state
    _nIdx    : INT;                        // 台索引 [-] / Stage index
    _nPick   : INT;                        // 候选台号 [-] / Candidate stage
    _bFound  : BOOL;                       // 候选已找到标志 [-] / Candidate found flag
    _bFault  : BOOL;                       // 故障锁存位（锁存量） / Latched fault bit
    _uFault  : UDINT;                      // 故障码锁存（锁存量） / Latched fault code
    _bCfgBad : BOOL;                       // 组态非法当拍量 [-] / Config illegal flag
    _bDemClp : BOOL;                       // 需量钳位当拍量 [-] / Demand clamped flag
    _bDwellLockCalc: BOOL;                 // 驻留阻塞内部量 [-] / Dwell blocking internal
    _uDwellOnScan: UDINT;                  // 运行驻留折算扫描数 [拍] / On dwell in scans
    _uDwellOffScan: UDINT;                 // 停机驻留折算扫描数 [拍] / Off dwell in scans
END_VAR
VAR CONSTANT
    DL_STAGE_MAX : INT := 4;               // 台数上限，与数组维度一致 [台] / Stage ceiling
    DL_ZERO_INT  : INT := 0;               // 零台常量 [台] / Zero stages
    DL_ZERO_UD   : UDINT := UDINT#0;       // 零计数常量 [拍] / Zero scans
    DL_MS_PER_MIN: REAL := 60000.0;        // 毫秒 → 分换算系数 [毫秒/分] / Milliseconds per minute
    DL_ONE_UD    : UDINT := UDINT#1;       // 单位计数常量 [拍] / One scan
END_VAR

(* —— 段 0｜沿与定时器每拍无条件刷新（禁置于 IF/CASE 内） —— *)
rtReset(CLK := bReset);
tonRotateWin(IN := (_eState = E_DL_CssState.eRun) AND (NOT _bFault) AND (NOT tonRotateWin.Q),
             PT := tRotateWin);          // 自复触周期窗：Q 拍断开一拍（R188）

(* —— 段 1｜瞬时量预清零（锁存量 _bFault/_uFault/abStageRun/auRunMin 不入清单） —— *)
uErrId   := 16#0000_0000;
_bCfgBad := FALSE;
_bDemClp := FALSE;

(* —— 段 2｜复位沿：故障一次性清干净，相位回空闲，全台停机 —— *)
IF rtReset.Q THEN
    _bFault := FALSE;
    _uFault := 16#0000_0000;
    FOR _nIdx := 1 TO DL_STAGE_MAX DO
        abStageRun[_nIdx] := FALSE;
        _abLastRun[_nIdx] := FALSE;
        _auDwellScan[_nIdx] := DL_ZERO_UD;
    END_FOR
    nStaged := DL_ZERO_INT;
    _eState := E_DL_CssState.eIdle;
END_IF

(* —— 段 3｜组态闸与需量钳位 —— *)
IF (tMinOn = T#0S) OR (tMinOff = T#0S) OR (tRotateWin = T#0S) OR (tCycle = T#0S) THEN
    _bCfgBad := TRUE;
END_IF
_nDemandUse := nDemand;
IF _nDemandUse < DL_ZERO_INT THEN
    _nDemandUse := DL_ZERO_INT;
    _bDemClp := TRUE;
ELSIF _nDemandUse > DL_STAGE_MAX THEN
    _nDemandUse := DL_STAGE_MAX;
    _bDemClp := TRUE;
END_IF
IF _bDemClp THEN
    uErrId := 16#0006_01BD;              // 信息级：需量钳位（瞬时口径）
END_IF

(* —— 段 4｜驻留折算：驻留时长 ÷ 扫描周期 = 驻留扫描数（除法前周期域闸已过） —— *)
_uDwellOnScan  := REAL_TO_UDINT(TIME_TO_REAL(tMinOn) / MAX(TIME_TO_REAL(tCycle), 1.0));
_uDwellOffScan := REAL_TO_UDINT(TIME_TO_REAL(tMinOff) / MAX(TIME_TO_REAL(tCycle), 1.0));

(* —— 段 5｜主状态机：三态全覆盖 + ELSE 兜底 —— *)
CASE _eState OF

E_DL_CssState.eIdle:
    FOR _nIdx := 1 TO DL_STAGE_MAX DO
        abStageRun[_nIdx] := FALSE;      // 空闲相全台停机（安全侧）
    END_FOR
    nStaged := DL_ZERO_INT;
    IF bEnable AND (NOT _bCfgBad) THEN
        FOR _nIdx := 1 TO DL_STAGE_MAX DO
            _auRunMin[_nIdx] := DL_ZERO_UD;      // 入运行相：运行时数基线清零
            _auDwellScan[_nIdx] := DL_ZERO_UD;
            _abLastRun[_nIdx] := FALSE;
        END_FOR
        _eState := E_DL_CssState.eRun;
    ELSIF bEnable AND _bCfgBad THEN
        _bFault := TRUE;
        _uFault := 16#0006_02BD;
        bError  := TRUE;
        _eState := E_DL_CssState.eFault;
    END_IF

E_DL_CssState.eRun:
    IF NOT bEnable THEN
        _eState := E_DL_CssState.eIdle;  // 使能撤销回空闲
    ELSE
        (* 运行时数与驻留计数：按上拍运行态刷新（驻留只在台数未变方向上累计） *)
        _bDwellLockCalc := FALSE;
        FOR _nIdx := 1 TO DL_STAGE_MAX DO
            IF abStageRun[_nIdx] THEN
                _auRunMin[_nIdx] := _auRunMin[_nIdx]
                    + REAL_TO_UDINT(TIME_TO_REAL(tCycle) / DL_MS_PER_MIN);
            END_IF
            IF abStageRun[_nIdx] = _abLastRun[_nIdx] THEN
                _auDwellScan[_nIdx] := _auDwellScan[_nIdx] + DL_ONE_UD;  // 方向未变：驻留累计
            ELSE
                _auDwellScan[_nIdx] := DL_ZERO_UD;   // 方向翻转：驻留清零
                _abLastRun[_nIdx] := abStageRun[_nIdx];
            END_IF
        END_FOR
        nStaged := DL_ZERO_INT;
        FOR _nIdx := 1 TO DL_STAGE_MAX DO
            IF abStageRun[_nIdx] THEN
                nStaged := nStaged + 1;
            END_IF
        END_FOR
        (* 加载：在编 < 需量，选运行时数最短的停机台（驻留满方可启） *)
        IF nStaged < _nDemandUse THEN
            _bFound := FALSE;
            _nPick  := 0;
            FOR _nIdx := 1 TO DL_STAGE_MAX DO
                IF (NOT abStageRun[_nIdx]) AND (_auDwellScan[_nIdx] >= _uDwellOffScan) THEN
                    IF (NOT _bFound) OR (_auRunMin[_nIdx] < _auRunMin[_nPick]) THEN
                        _bFound := TRUE;
                        _nPick  := _nIdx;
                    END_IF
                END_IF
            END_FOR
            IF _bFound THEN
                abStageRun[_nPick] := TRUE;  // 启动轮值均衡最优台
                _abLastRun[_nPick] := TRUE;
                _auDwellScan[_nPick] := DL_ZERO_UD;
            ELSE
                _bDwellLockCalc := TRUE;     // 无驻留满足台：阻塞
            END_IF
        ELSIF nStaged > _nDemandUse THEN
            (* 卸载：在编 > 需量，选运行时数最长的运行台（驻留满方可停） *)
            _bFound := FALSE;
            _nPick  := 0;
            FOR _nIdx := 1 TO DL_STAGE_MAX DO
                IF abStageRun[_nIdx] AND (_auDwellScan[_nIdx] >= _uDwellOnScan) THEN
                    IF (NOT _bFound) OR (_auRunMin[_nIdx] > _auRunMin[_nPick]) THEN
                        _bFound := TRUE;
                        _nPick  := _nIdx;
                    END_IF
                END_IF
            END_FOR
            IF _bFound THEN
                abStageRun[_nPick] := FALSE; // 停止轮值均衡最劣台
                _abLastRun[_nPick] := FALSE;
                _auDwellScan[_nPick] := DL_ZERO_UD;
            ELSE
                _bDwellLockCalc := TRUE;     // 无驻留满足台：阻塞
            END_IF
        END_IF
        bDwellLock := _bDwellLockCalc;       // 驻留阻塞电平同源赋值（R191）
    END_IF

E_DL_CssState.eFault:
    FOR _nIdx := 1 TO DL_STAGE_MAX DO
        abStageRun[_nIdx] := FALSE;      // 故障相全台停机（安全侧）
    END_FOR
    nStaged := DL_ZERO_INT;
    bError := TRUE;
    ;                                    // 故障相驻留：只认复位沿（段 2 迁出）

ELSE
    _bFault := TRUE;                     // 兜底：非法相位锁存
    _uFault := 16#0006_02BD;
    bError  := TRUE;
    _eState := E_DL_CssState.eFault;
END_CASE

(* —— 段 6｜状态出口单点映射 —— *)
eState := _eState;
END_FUNCTION_BLOCK

(* ---- FB_DL_ChillerTempStab.st ---- *)
(*==============================================================================
 * 组件名称 (Component)  : FB_DL_ChillerTempStab
 * 溯源说明 (Provenance) : 道莅 clean-room 防御性实现（路线图 L259 已登记项）
 * 所属子库 (Sublibrary) : DL_Process / ProcessStability
 * 当前版本 (Version)    : 1.0.0
 * 兼容性   (Platform)   : CODESYS 3.5 / TwinCAT 3 / 汇川 InoProShop；
 *                         纯 IEC 61131-3（第 3 版），仅用标准库 TON
 * 组件分类 (Category)   : 功能块（FUNCTION_BLOCK）· 冷冻水供水温度稳定性监视
 * 功能一句话 (Summary)  : 双代滑窗均值/标准差 + CV 判稳 + 不稳定确认延时。
 * 边界与安全 (Boundary) : ①温度 NaN 或超出 -40~120 ℃ 拒收并置码；
 *                         ②样本数不足最小值 → bStable=FALSE 且不判稳；
 *                         ③均值绝对值近零时 CV 分母防御（除零前判）；
 *                         ④不稳定确认 TON 无条件周期刷新；
 *                         ⑤bReset 清全部统计（重新起窗）。
 * 错误码    : 16#0005_035F 样本非法拒收（NaN 或超量程）——故障级（持续态）
 *             16#0005_0360 判稳确认超时未达成（持续不稳）——故障级（持续态）
 * 码位总账  : 16#0005_035F 用 / 16#0005_0360 用
 * 修改记录  : v1.0.0 R26 初版
 *==============================================================================*)
FUNCTION_BLOCK FB_DL_ChillerTempStab
VAR_INPUT
    fSupplyTemp : LREAL; // 供水温度 [℃] / Supply water temperature [degC]
    fCvLimit    : LREAL; // 变异系数判稳门限 [%] / CV stability limit [%]
    tConfirm    : TIME;  // 不稳定确认延时 [ms] / Instability confirm delay [ms]
    bReset      : BOOL;  // 复位：清统计重起窗 / Reset: clear statistics
    bEnable     : BOOL;  // 监视使能 / Monitoring enable
END_VAR
VAR_OUTPUT
    fMean            : LREAL; // 滑窗均值 [℃] / Sliding window mean [degC]
    fStdDev          : LREAL; // 滑窗标准差 [℃] / Sliding window std-dev [degC]
    fCv              : LREAL; // 变异系数 [%] / Coefficient of variation [%]
    bStable          : BOOL;  // 判稳结论 / Stability verdict
    bUnstableConfirm : BOOL;  // 不稳定确认（延时满足）/ Instability confirmed
    eErr             : UDINT; // 本周期错误码，0=无错 / Error code this cycle, 0 = none
END_VAR
VAR CONSTANT
    cHalves  : DINT  := 10;    // 窗内代数（双代近似滑窗）/ Window generations
    cMinSmp  : UDINT := 30;    // 最小样本数 / Minimum sample count
    cTempLo  : LREAL := -40.0; // 温度下限 [℃] / Temperature lower bound
    cTempHi  : LREAL := 120.0; // 温度上限 [℃] / Temperature upper bound
END_VAR
VAR
    fSumOld : LREAL; // 旧代样本和 / Previous generation sum
    fSqOld  : LREAL; // 旧代平方和 / Previous generation sum of squares
    fSumNew : LREAL; // 新代样本和 / Current generation sum
    fSqNew  : LREAL; // 新代平方和 / Current generation sum of squares
    uCntOld : UDINT; // 旧代样本数 / Previous generation count
    uCntNew : UDINT; // 新代样本数 / Current generation count
    iGen    : INT;   // 当前代序号 / Current generation index
    tonGen  : TON;   // 代轮转定时器（无条件刷新）/ Generation rotation timer
    tonUnst : TON;   // 不稳定确认定时器（无条件刷新）/ Instability confirm timer
    dwGenMs : DINT;  // 单代时长 [ms] / Generation duration [ms]
    fVarAll : LREAL; // 总体方差临时量 / Total variance temp
    bSmpOk  : BOOL;  // 本拍样本合法性 / Sample validity this cycle
END_VAR

// ---------- 代时长：确认窗 / 代数（下限防御） ----------
dwGenMs := TIME_TO_DINT(tConfirm) / cHalves;
IF dwGenMs < 1 THEN
    dwGenMs := 1;                             // 最小 1 ms 代 / Minimum 1 ms generation
END_IF
tonGen(IN := bEnable, PT := DINT_TO_TIME(dwGenMs));

// ---------- 复位与禁能清统计 ----------
IF bReset OR (NOT bEnable) THEN
    fSumOld := 0.0; fSqOld := 0.0; fSumNew := 0.0; fSqNew := 0.0;
    uCntOld := 0;   uCntNew := 0;  iGen := 0;
    fMean := 0.0; fStdDev := 0.0; fCv := 0.0;
    bStable := FALSE;
    bUnstableConfirm := FALSE;
END_IF

// ---------- 样本防御：NaN 或超量程拒收 ----------
bSmpOk := FALSE;
IF bEnable THEN
    eErr := 0;
    IF (fSupplyTemp <> fSupplyTemp) OR ((fSupplyTemp - fSupplyTemp) <> (fSupplyTemp - fSupplyTemp)) THEN
        eErr := 16#0005_035F;                 // NaN 拒收 / NaN rejected
    ELSIF (fSupplyTemp < cTempLo) OR (fSupplyTemp > cTempHi) THEN
        eErr := 16#0005_035F;                 // 超量程拒收 / Out-of-range rejected
    ELSE
        bSmpOk := TRUE;                       // 合法样本 / Valid sample
    END_IF
END_IF

// ---------- 合法样本入新代 ----------
IF bSmpOk THEN
    fSumNew := fSumNew + fSupplyTemp;         // 样本和 / Sample sum
    fSqNew  := fSqNew + fSupplyTemp * fSupplyTemp; // 平方和 / Square sum
    uCntNew := uCntNew + UDINT#1;             // 计数 / Count
END_IF

// ---------- 代轮转（与扭矩监视件同口径双代近似） ----------
IF tonGen.Q THEN
    iGen := iGen + 1;
    IF iGen >= cHalves THEN
        iGen := cHalves / 2;
        fSumOld := fSumNew; fSqOld := fSqNew; uCntOld := uCntNew; // 新代平移 / Shift
        fSumNew := 0.0; fSqNew := 0.0; uCntNew := 0;              // 新代清零 / Clear
    END_IF
END_IF

// ---------- 均值/标准差/CV 计算（除法全部前判零） ----------
IF (uCntOld + uCntNew) >= cMinSmp THEN
    fMean := (fSumOld + fSumNew) / UDINT_TO_LREAL(uCntOld + uCntNew);   // 均值 / Mean
    fVarAll := (fSqOld + fSqNew) / UDINT_TO_LREAL(uCntOld + uCntNew) - fMean * fMean; // 方差 / Variance
    IF fVarAll < 0.0 THEN
        fVarAll := 0.0;                       // 数值误差负方差钳零 / Clamp tiny negative variance
    END_IF
    fStdDev := SQRT(fVarAll);                 // 标准差 / Std-dev
    IF ABS(fMean) > 1.0E-9 THEN
        fCv := fStdDev / ABS(fMean) * 100.0;  // 变异系数 / CV in percent
    ELSE
        fCv := 0.0;                           // 近零均值 CV 防御 / Near-zero mean guard
    END_IF
    bStable := fCv <= fCvLimit;               // 判稳结论 / Stability verdict
ELSE
    fMean := 0.0;                             // 样本不足不出值 / Insufficient samples
    fStdDev := 0.0;
    fCv := 0.0;
    bStable := FALSE;                         // 未满窗不判稳 / No verdict before window filled
END_IF

// ---------- 无条件周期刷新：不稳定确认定时器 ----------
tonUnst(IN := bEnable AND (NOT bStable), PT := tConfirm);
IF tonUnst.Q THEN
    bUnstableConfirm := TRUE;                 // 确认成立 / Confirmed
    eErr := 16#0005_0360;                     // 判稳超时未达成码 / Never-stable confirm code
ELSE
    bUnstableConfirm := FALSE;                // 未确认即撤销 / Withdrawn if unconfirmed
END_IF

END_FUNCTION_BLOCK
